(* IEC 61131-3 sources: daoli-st-library/DL_Algo (part 16) *)

(* ---- FB_DL_LoopCoupleDetect.st ---- *)
(*==============================================================================
 * 组件名称 (Component)  : FB_DL_LoopCoupleDetect
 * 所属子库 (Sublibrary) : DL_Algo
 * 当前版本 (Version)    : 1.0.1
 * 兼容性 (Platform)     : CODESYS 3.5+ / TwinCAT 3 / 汇川 InoProShop / 施耐德 Machine Expert
 *                         仅依赖 Standard.library（TON / R_TRIG），零厂商私有库
 * 功能描述 (Function)   : 回路耦合度在线探测。本回路上位激励期（bExcite 电平）
 *                         同步采集本回路 CV 增量 x 与邻回路 PV 增量 y，窗口内
 *                         计算皮尔逊互相关系数 r；|r| >= fCoupleThresh 且样本
 *                         充分 → bCoupled 锁存并输出耦合强度分级。为 Decouple2x2
 *                         提供投运判据（探测在先、解耦执行在后）。
 * 来源标签 (Origin)     : 自研线（IEC 61131-3 标准语义的道莅防御性实现，clean-room）
 * 分工声明 (Pairing)    : LoopCoupleDetect（探测，本件）↔ FB_DL_Decouple2x2
 *                         （解耦执行，既有件）：本件只输出耦合判据与强度分级，
 *                         不注入任何解耦补偿量、不修改解耦矩阵（R298 属主边界）；
 *                         与 FB_DL_CrossCorrelationDelay 分工：本件测「响应强度」
 *                         不测「延时幅值」，二者互补不重叠。
 * 边界语义 (Boundary)   : ① 相关系数除零防御：任一分母因子 <= eps → r 按 0
 *                         （邻回路无响应 = 无耦合语义，合法结果非故障）；
 *                         ② 非激励期（bExcite = FALSE）不采样不判据（判据串
 *                         相位因子，R281 口径）；
 *                         ③ 增量非有限拒收（NaN 自反 + Inf 差判）；
 *                         ④ 组态闸：窗深/阈值/最小样本 → 故障锁存。
 * 输出语义 (Fallback)   : 【R191】非激励期 → fCorrOut 保持末值、bCoupled 保持
 *                         锁存（耦合是资产属性，不随激励停而消失）；eFault 相
 *                         → 冻结 + bError = TRUE。
 * 码位     (Codes)      : 按 R297 范式零 16# 码位硬编码；错误出口 BOOL+ENUM(eCause)，
 *                         码位待主控收口统一派号。
 * 红线自检 (Redline)    : 7 项红线已自检：R1 零全局 ✓｜R2 零物理地址 ✓｜R3 纯 IEC ✓
 *                         R4 除零（双因子 eps 闸）/NaN 拒收/组态闸 ✓
 *                         R5 双语同行注释 ✓｜R6 CASE 带 ELSE 兜底迁 eFault ✓
 *                         R7 TON/R_TRIG 段 0 无条件刷新 ✓
 * 验收向量 (Acceptance) : V1 强耦合仿真（y = 0.8·x + 噪声）→ |r| ≈ 0.8+，
 *                         eStrength=eStrong，bCoupled=TRUE；
 *                         V2 独立回路（y 与 x 无关）→ |r| < 阈值，
 *                         eStrength=eNone；
 *                         V3 非激励期停止采样，样本数不增。
 * 修订历史 (Revision)   : 2026-11-20  v1.0.0  R49 首版（批 3 · 序号 13）
 *                        2026-11-20  v1.0.1  R51 文档级更正（R50 终审轻项）：3 处
 *                        相对指代禁词注释改为自含描述（R92/R68）；逻辑零变更
 *==============================================================================*)
TYPE E_DL_LcdStrength :
(
    eNone    := 0,                           (* 无耦合：|r| < 弱阈值 / No coupling *)
    eWeak    := 1,                           (* 弱耦合：|r| ∈ [弱阈, 强阈) / Weak coupling *)
    eStrong  := 2                            (* 强耦合：|r| >= 强阈值 / Strong coupling *)
);
END_TYPE

TYPE E_DL_LcdState :
(
    eIdle  := 0,                             (* 待使能 / Idle *)
    eProbe := 10,                            (* 激励探测运行 / Excitation probing *)
    eFault := 90                             (* 故障锁存相 / Fault latched phase *)
);
END_TYPE

TYPE E_DL_LcdCause :
(
    eNone       := 0,                        (* 无故障成因 / No cause *)
    eCfgIllegal := 1,                        (* 组态非法：窗深/阈值越域 / Illegal config *)
    ePhaseBad   := 2                         (* 非法相位兜底 / Illegal phase fallback *)
);
END_TYPE

FUNCTION_BLOCK FB_DL_LoopCoupleDetect
VAR_INPUT
    fCvThis   : LREAL := 0.0;                (* 本回路 CV 当前值（激励侧）[工程单位] / This loop CV value *)
    fPvNeighbor : LREAL := 0.0;              (* 邻回路 PV 当前值（响应侧）[工程单位] / Neighbor loop PV value *)
    bExcite   : BOOL := FALSE;               (* 本回路激励期电平（上位投运流程给出）[-] / Excitation period level *)
    nWinDepth : INT := 64;                   (* 互相关窗深，域 8..128 [点] / Correlation window depth *)
    fCoupleThresh : LREAL := 0.5;            (* 耦合判据阈值（|r| 门限），域 (0,1) [-] / Coupling threshold *)
    bEnable   : BOOL := TRUE;                (* 探测使能 [-] / Enable *)
    bReset    : BOOL := FALSE;               (* 复位命令，上升沿清窗与全部锁存 [-] / Reset command *)
END_VAR
VAR_OUTPUT
    fCorrOut  : LREAL;                       (* 当前窗口互相关系数 [-] / Window correlation coefficient *)
    eStrength : E_DL_LcdStrength;            (* 耦合强度分级出口（按最新窗口派生）[-] / Coupling strength outlet *)
    bCoupled  : BOOL;                        (* 耦合判据锁存位（复位沿清）[-] / Coupled latch *)
    nSampleCnt: INT;                         (* 窗口有效样本数 [点] / Valid sample count *)
    eState    : E_DL_LcdState;               (* 状态出口 / State outlet *)
    eCause    : E_DL_LcdCause;               (* 故障成因出口（R190 归因唯一） / Fault cause outlet *)
    bError    : BOOL;                        (* 故障锁存标志 [-] / Fault latch flag *)
END_VAR
VAR
    _eState  : E_DL_LcdState := E_DL_LcdState.eIdle;      (* 内部相位（CASE 唯一写入目标） / Internal phase *)
    _eCause  : E_DL_LcdCause := E_DL_LcdCause.eNone;      (* 故障成因锁存量 / Latched cause *)
    rtReset  : R_TRIG;                       (* 复位沿实例，段 0 无条件调用 / Reset edge instance *)
    _fCvPrev : LREAL;                        (* 上拍本回路 CV（增量基准）[工程单位] / Previous this-loop CV *)
    _fPvPrev : LREAL;                        (* 上拍邻回路 PV（增量基准）[工程单位] / Previous neighbor PV *)
    _aDx     : ARRAY[1..128] OF LREAL;       (* 本回路 CV 增量窗 [工程单位] / This-loop dCV window *)
    _aDy     : ARRAY[1..128] OF LREAL;       (* 邻回路 PV 增量窗 [工程单位] / Neighbor dPV window *)
    _nHead   : INT;                          (* 环形头游标 [-] / Ring head cursor *)
    _nFill   : INT;                          (* 窗填充数 [点] / Window fill count *)
    _nEff    : INT;                          (* 钳位后生效窗深 [点] / Clamped effective depth *)
    _fSumX   : LREAL;                        (* Σx [工程单位] / Sum x *)
    _fSumY   : LREAL;                        (* Σy [工程单位] / Sum y *)
    _fSumXY  : LREAL;                        (* Σxy [工程单位²] / Sum xy *)
    _fSumX2  : LREAL;                        (* Σx² [工程单位²] / Sum x2 *)
    _fSumY2  : LREAL;                        (* Σy² [工程单位²] / Sum y2 *)
    _fDen    : LREAL;                        (* 分母乘积（开方前）[-] / Denominator product *)
    _fR      : LREAL;                        (* 本拍相关系数 [-] / Correlation this scan *)
    _bFault  : BOOL;                         (* 故障锁存位 / Latched fault bit *)
    _bCfgBad : BOOL;                         (* 组态非法当拍量 / Illegal config this scan *)
    _i       : INT;                          (* 统计扫描游标（每趟重置，R227）[-] / Stats cursor *)
END_VAR
VAR CONSTANT
    DL_LCD_EPS  : LREAL := 1.0E-12;          (* 分母因子判零容差 [-] / Denominator epsilon *)
    DL_LCD_NMAX : INT   := 128;              (* 窗深容量上限 [点] / Window capacity limit *)
    DL_LCD_MIN  : INT   := 16;               (* 判据最小样本数（不足不判，防短窗误报）[点] / Min samples for verdict *)
    DL_LCD_WEAK : LREAL := 0.3;              (* 弱耦合门限（强度分级内界）[-] / Weak coupling bound *)
END_VAR

(* —— 段 0：当拍判据派生 + 实例无条件刷新（R228A） —— *)
_bCfgBad := (nWinDepth < 8) OR (nWinDepth > DL_LCD_NMAX) OR (fCoupleThresh <= 0.0) OR (fCoupleThresh >= 1.0);   (* 组态闸（R151 全引脚） / Config gate *)
rtReset(CLK := bReset);                      (* 复位沿每拍必调 / Reset edge every scan *)
_nEff := nWinDepth;                          (* 生效窗深初值 / Depth init *)
IF _nEff < 8 THEN
    _nEff := 8;                              (* 下限钳位 / Lower clamp *)
END_IF
IF _nEff > DL_LCD_NMAX THEN
    _nEff := DL_LCD_NMAX;                    (* 上限钳位（R308） / Upper clamp *)
END_IF

(* —— 段 1：单拍量预清零（R107） —— *)
_fSumX := 0.0;                               (* 累计量清零重算（每拍全路径派生，R285） / Sums recompute *)
_fSumY := 0.0;                               (* Σy 清零 / Sum y clear *)
_fSumXY := 0.0;                              (* Σxy 清零 / Sum xy clear *)
_fSumX2 := 0.0;                              (* Σx² 清零 / Sum x2 clear *)
_fSumY2 := 0.0;                              (* Σy² 清零 / Sum y2 clear *)
_fDen := 0.0;                                (* 分母清零（防残留触发除零） / Denominator clear *)
_fR := 0.0;                                  (* 相关系数缺省 0 / Correlation default *)

(* —— 段 2：复位沿处理（作用域：清故障 + 清窗 + 清锁存 + 基准重锚 + 迁 eIdle，R283 逐项声明） —— *)
IF rtReset.Q THEN
    _bFault := FALSE;                        (* 清故障锁存 / Clear fault *)
    _eCause := E_DL_LcdCause.eNone;          (* 清成因 / Clear cause *)
    _nFill := 0;                             (* 清窗填充 / Clear fill *)
    _nHead := 1;                             (* 头游标复位 / Head reset *)
    bCoupled := FALSE;                       (* 清耦合锁存 / Clear coupled latch *)
    fCorrOut := 0.0;                         (* 清相关系数出口 / Clear correlation outlet *)
    _fCvPrev := fCvThis;                     (* 增量基准重锚 / Re-anchor base *)
    _fPvPrev := fPvNeighbor;                 (* 邻回路 PV 增量基准重锚 / Re-anchor neighbor PV base *)
    _eState := E_DL_LcdState.eIdle;          (* 迁待机相 / Back to idle *)
END_IF

(* —— 段 3：组态闸故障锁存（R45 配对；锁存至复位沿，R189） —— *)
IF _bCfgBad AND NOT _bFault THEN
    _bFault := TRUE;                         (* 锁存故障位 / Latch fault *)
    _eCause := E_DL_LcdCause.eCfgIllegal;    (* 成因：组态非法 / Cause: illegal config *)
    _eState := E_DL_LcdState.eFault;         (* 同步迁故障相 / Migrate to fault *)
END_IF

(* —— 段 4：CASE 主状态机（ELSE 兜底迁 eFault，红线 6） —— *)
CASE _eState OF
    E_DL_LcdState.eIdle:                     (* 待机相：基准持续跟锚 / Idle *)
        _fCvPrev := fCvThis;                 (* 防待机期巨增量 / Anchor follow *)
        _fPvPrev := fPvNeighbor;             (* 邻回路 PV 基准持续跟锚（防待机期巨增量） / Neighbor PV base follow *)
        IF bEnable AND NOT _bFault THEN
            _eState := E_DL_LcdState.eProbe; (* 进入探测 / Enter probe *)
        END_IF
    E_DL_LcdState.eProbe:                    (* 探测相：仅激励期采样 + 窗口统计 / Probe *)
        IF NOT bEnable THEN
            _eState := E_DL_LcdState.eIdle;  (* 失能回待机 / Back to idle *)
        ELSE
            IF bExcite THEN                  (* 判据串相位因子：仅激励期采样（R281） / Sample only in excitation *)
                _aDx[_nHead] := fCvThis - _fCvPrev;       (* 本回路 CV 增量入窗 / This-loop dCV *)
                _aDy[_nHead] := fPvNeighbor - _fPvPrev;   (* 邻回路 PV 增量入窗 / Neighbor dPV *)
                IF (_aDx[_nHead] <> _aDx[_nHead]) OR (_aDy[_nHead] <> _aDy[_nHead])
                   OR ((_aDx[_nHead] - _aDx[_nHead]) <> (_aDx[_nHead] - _aDx[_nHead]))
                   OR ((_aDy[_nHead] - _aDy[_nHead]) <> (_aDy[_nHead] - _aDy[_nHead])) THEN
                    (* 非有限增量：不入统计不推进游标，基准照常跟锚 / Non-finite: skip *)
                    ;                        (* 空语句：ST 语法要求 THEN 分支非空，无副作用 / Empty statement, ST syntax requires non-empty branch *)
                ELSE
                    _nHead := _nHead + 1;    (* 有效样本：游标递进 / Head advance *)
                    IF _nHead > _nEff THEN
                        _nHead := 1;         (* 环回卷 / Ring wrap *)
                    END_IF
                    IF _nFill < _nEff THEN
                        _nFill := _nFill + 1;    (* 填充封顶 / Fill cap *)
                    END_IF
                END_IF
                _fCvPrev := fCvThis;         (* 基准推进 / Base advance *)
                _fPvPrev := fPvNeighbor;     (* 邻回路 PV 基准推进（与本拍采样配对） / Neighbor PV base advance *)
            END_IF
            _i := 1;                         (* 统计游标起头重置（R227） / Cursor reset *)
            WHILE _i <= _nFill DO            (* 逐点累计 / Per-point sums *)
                _fSumX := _fSumX + _aDx[_i]; (* Σx / Sum x *)
                _fSumY := _fSumY + _aDy[_i]; (* Σy / Sum y *)
                _fSumXY := _fSumXY + _aDx[_i] * _aDy[_i];   (* Σxy / Sum xy *)
                _fSumX2 := _fSumX2 + _aDx[_i] * _aDx[_i];   (* Σx² / Sum x2 *)
                _fSumY2 := _fSumY2 + _aDy[_i] * _aDy[_i];   (* Σy² / Sum y2 *)
                _i := _i + 1;                (* 游标递进 / Cursor advance *)
            END_WHILE
            IF _nFill >= 1 THEN
                _fDen := (DINT_TO_LREAL(_nFill) * _fSumX2 - _fSumX * _fSumX)
                       * (DINT_TO_LREAL(_nFill) * _fSumY2 - _fSumY * _fSumY);   (* 分母乘积（双因子联合闸） / Denominator product *)
            END_IF
            IF (_fDen > DL_LCD_EPS * DL_LCD_EPS) AND (_nFill >= 1) THEN
                _fR := (DINT_TO_LREAL(_nFill) * _fSumXY - _fSumX * _fSumY) / SQRT(_fDen);   (* 互相关 r：分母已过联合 eps 闸，无除零 / Correlation, denominator gated *)
                fCorrOut := _fR;             (* 相关系数出口更新（仅有效窗刷新） / Update outlet *)
                IF (_nFill >= DL_LCD_MIN) AND (_nFill * 10 >= 6 * _nEff) THEN
                    IF ABS(_fR) >= fCoupleThresh THEN
                        bCoupled := TRUE;    (* 耦合判据锁存至复位沿 / Coupled latch *)
                    END_IF
                    IF ABS(_fR) >= fCoupleThresh THEN
                        eStrength := E_DL_LcdStrength.eStrong;   (* 强耦合 / Strong *)
                    ELSIF ABS(_fR) >= DL_LCD_WEAK THEN
                        eStrength := E_DL_LcdStrength.eWeak;     (* 弱耦合 / Weak *)
                    ELSE
                        eStrength := E_DL_LcdStrength.eNone;     (* 无耦合（IF 链带 ELSE 兜底，R285） / None *)
                    END_IF
                END_IF
            END_IF
            nSampleCnt := _nFill;            (* 样本数出口镜像 / Sample count mirror *)
        END_IF
    E_DL_LcdState.eFault:                    (* 故障相：冻结保持，仅复位沿出 / Fault *)
        ;                                    (* 锁存回放（R28） / Replay from latch *)
    ELSE                                     (* 非法相位兜底迁安全态 / Illegal phase fallback *)
        _eState := E_DL_LcdState.eFault;     (* 迁故障相 / To fault *)
        _bFault := TRUE;                     (* 同步锁存 / Latch *)
        _eCause := E_DL_LcdCause.ePhaseBad;  (* 成因：非法相位 / Cause: illegal phase *)
END_CASE

(* —— 段 5：出口映射（bError/eState 同源，R191） —— *)
bError := _bFault;                           (* 故障标志镜像 / Fault flag mirror *)
eState := _eState;                           (* 状态出口 / State outlet *)
eCause := _eCause;                           (* 成因出口 / Cause outlet *)
END_FUNCTION_BLOCK

(* ---- FB_DL_LoopSignGuard.st ---- *)
(*==============================================================================
 * 组件名称 (Component)  : FB_DL_LoopSignGuard
 * 所属子库 (Sublibrary) : DL_Algo
 * 当前版本 (Version)    : 1.0.0
 * 兼容性 (Platform)     : CODESYS 3.5+ / TwinCAT 3 / 汇川 InoProShop / 施耐德 Machine Expert
 *                         仅依赖 Standard.library（TON），零厂商私有库
 * 功能描述 (Function)   : 回路正反作用符号在线自检（调试期防呆）。以增量对
 *                         (dCV, dPV) 为样本，窗口内计算皮尔逊相关系数
 *                         r = (nΣxy - ΣxΣy) / sqrt((nΣx²-(Σx)²)·(nΣy²-(Σy)²))：
 *                         r > fSignThresh → 判正向作用（CV 增大 PV 随之增大）；
 *                         r < -fSignThresh → 判反向作用；|r| 不足 → 未定。
 *                         期望作用 eExpect 与实测作用不一致 → bSignSuspect
 *                         锁存（接线反接/正反作用组态错防呆）。
 * 来源标签 (Origin)     : 自研线（IEC 61131-3 标准语义的道莅防御性实现，clean-room）
 * 边界语义 (Boundary)   : ① 相关系数除零防御：分母任一因子 <= eps（窗口内
 *                         CV 或 PV 无变化，如手动手假输入）→ r 按 0 处理（未定），
 *                         不产生 Inf/NaN；
 *                         ② 样本拒收：dCV/dPV 非有限（NaN/Inf 差判）不入窗；
 *                         ③ 判据串相位因子：仅 nSample >= 窗深 60% 后才判
 *                         （样本不足不判，防启动段误报，R281 口径）；
 *                         ④ 组态闸：窗深 < 8 / 阈值域 (0,1) 外 → 故障。
 * 输出语义 (Fallback)   : 【R191】样本不足期 → eSignOut = eUnknown，bSignSuspect
 *                         保持 FALSE；eFault 相 → 判据输出冻结保持末值。
 * 码位     (Codes)      : 按 R297 范式零 16# 码位硬编码；错误出口 BOOL+ENUM(eCause)，
 *                         码位待主控收口统一派号。
 * 红线自检 (Redline)    : 7 项红线已自检：R1 零全局 ✓｜R2 零物理地址 ✓｜R3 纯 IEC ✓
 *                         R4 除零（双因子 eps 闸）/NaN 拒收/组态闸 ✓
 *                         R5 双语同行注释 ✓｜R6 CASE 带 ELSE 兜底迁 eFault ✓
 *                         R7 TON/R_TRIG 段 0 无条件刷新 ✓
 * 验收向量 (Acceptance) : V1 同向增量样本 32 点 → r≈1 → eSignOut=eDirect；
 *                         V2 反向增量样本 → r≈-1 → eSignOut=eReverse，若
 *                         eExpect=eDirect → bSignSuspect=TRUE；
 *                         V3 恒定 PV（分母 0）→ eSignOut=eUnknown，不误报。
 * 修订历史 (Revision)   : 2026-11-20  v1.0.0  R49 首版（批 3 · 序号 11）
 *==============================================================================*)
TYPE E_DL_LsgSign :
(
    eUnknown := 0,                           (* 未定（样本不足或相关性弱） / Unknown *)
    eDirect  := 1,                           (* 正向作用：CV↑ → PV↑ / Direct acting *)
    eReverse := 2                            (* 反向作用：CV↑ → PV↓ / Reverse acting *)
);
END_TYPE

TYPE E_DL_LsgState :
(
    eIdle  := 0,                             (* 待使能 / Idle *)
    eLearn := 10,                            (* 增量样本采集学习中 / Learning *)
    eFault := 90                             (* 故障锁存相 / Fault latched phase *)
);
END_TYPE

TYPE E_DL_LsgCause :
(
    eNone       := 0,                        (* 无故障成因 / No cause *)
    eCfgIllegal := 1,                        (* 组态非法：窗深/阈值越域 / Illegal config *)
    ePhaseBad   := 2                         (* 非法相位兜底 / Illegal phase fallback *)
);
END_TYPE

FUNCTION_BLOCK FB_DL_LoopSignGuard
VAR_INPUT
    fCvNow    : LREAL := 0.0;                (* 控制量当前值（CV）[工程单位] / CV current value *)
    fPvNow    : LREAL := 0.0;                (* 过程量当前值（PV）[工程单位] / PV current value *)
    nWinDepth : INT := 32;                   (* 增量样本窗深，域 8..64 [点] / Sample window depth *)
    fSignThresh : LREAL := 0.6;              (* 判向阈值（|r| 门限），域 (0.0, 1.0) [-] / Sign verdict threshold *)
    eExpect   : E_DL_LsgSign := E_DL_LsgSign.eDirect;   (* 期望作用方向（组态声明）[-] / Expected acting direction *)
    bEnable   : BOOL := TRUE;                (* 自检使能 [-] / Enable *)
    bReset    : BOOL := FALSE;               (* 复位命令，上升沿清全部样本与锁存 [-] / Reset command *)
END_VAR
VAR_OUTPUT
    eSignOut     : E_DL_LsgSign;             (* 实测作用方向出口 / Measured sign outlet *)
    fCorrCoef    : LREAL;                    (* 当前窗口皮尔逊相关系数 [-] / Pearson correlation of window *)
    nSampleCnt   : INT;                      (* 窗口内有效样本数 [点] / Valid sample count *)
    bSignSuspect : BOOL;                     (* 作用方向与期望不符锁存位（复位沿清）[-] / Sign-suspect latch *)
    eState       : E_DL_LsgState;            (* 状态出口 / State outlet *)
    eCause       : E_DL_LsgCause;            (* 故障成因出口（R190 归因唯一） / Fault cause outlet *)
    bError       : BOOL;                     (* 故障锁存标志 [-] / Fault latch flag *)
END_VAR
VAR
    _eState  : E_DL_LsgState := E_DL_LsgState.eIdle;      (* 内部相位（CASE 唯一写入目标） / Internal phase *)
    _eCause  : E_DL_LsgCause := E_DL_LsgCause.eNone;      (* 故障成因锁存量 / Latched cause *)
    rtReset  : R_TRIG;                       (* 复位沿实例，段 0 无条件调用 / Reset edge instance *)
    _fCvPrev : LREAL;                        (* 上拍 CV（增量基准）[工程单位] / Previous CV *)
    _fPvPrev : LREAL;                        (* 上拍 PV（增量基准）[工程单位] / Previous PV *)
    _aDx     : ARRAY[1..64] OF LREAL;        (* dCV 样本窗 [工程单位] / dCV window *)
    _aDy     : ARRAY[1..64] OF LREAL;        (* dPV 样本窗 [工程单位] / dPV window *)
    _nHead   : INT;                          (* 环形头游标 [-] / Ring head cursor *)
    _nFill   : INT;                          (* 窗口填充数 [点] / Window fill count *)
    _nEff    : INT;                          (* 钳位后生效窗深 [点] / Clamped effective depth *)
    _fSumX   : LREAL;                        (* Σx 累计 [工程单位] / Sum x *)
    _fSumY   : LREAL;                        (* Σy 累计 [工程单位] / Sum y *)
    _fSumXY  : LREAL;                        (* Σxy 累计 [工程单位²] / Sum xy *)
    _fSumX2  : LREAL;                        (* Σx² 累计 [工程单位²] / Sum x2 *)
    _fSumY2  : LREAL;                        (* Σy² 累计 [工程单位²] / Sum y2 *)
    _fDenX   : LREAL;                        (* 分母因子 1：nΣx²-(Σx)² [-] / Denominator factor 1 *)
    _fDenY   : LREAL;                        (* 分母因子 2：nΣy²-(Σy)² [-] / Denominator factor 2 *)
    _fDen    : LREAL;                        (* 相关系数分母（开方前乘积）[-] / Correlation denominator *)
    _fR      : LREAL;                        (* 本拍相关系数 [-] / Correlation this scan *)
    _eSign   : E_DL_LsgSign := E_DL_LsgSign.eUnknown;     (* 实测方向锁存 / Measured sign latch *)
    _bFault  : BOOL;                         (* 故障锁存位 / Latched fault bit *)
    _bCfgBad : BOOL;                         (* 组态非法当拍量 / Illegal config this scan *)
    _i       : INT;                          (* 统计扫描游标（每趟重置，R227）[-] / Stats cursor *)
END_VAR
VAR CONSTANT
    DL_LSG_EPS   : LREAL := 1.0E-12;         (* 分母因子判零容差 [-] / Denominator epsilon *)
    DL_LSG_NMAX  : INT   := 64;              (* 窗深容量上限 [点] / Window capacity limit *)
END_VAR

(* —— 段 0：当拍判据派生 + 实例无条件刷新（R228A） —— *)
_bCfgBad := (nWinDepth < 8) OR (nWinDepth > DL_LSG_NMAX) OR (fSignThresh <= 0.0) OR (fSignThresh >= 1.0);   (* 组态闸（R151 全引脚） / Config gate *)
rtReset(CLK := bReset);                      (* 复位沿每拍必调 / Reset edge every scan *)
_nEff := nWinDepth;                          (* 生效窗深初值 / Effective depth init *)
IF _nEff < 8 THEN
    _nEff := 8;                              (* 窗深下限钳位 / Depth lower clamp *)
END_IF
IF _nEff > DL_LSG_NMAX THEN
    _nEff := DL_LSG_NMAX;                    (* 窗深上限钳位（R308） / Depth upper clamp *)
END_IF

(* —— 段 1：单拍量预清零（R107） —— *)
_fSumX := 0.0;                               (* 累计量清零重算（每拍全路径派生，R285） / Sums recompute *)
_fSumY := 0.0;                               (* Σy 清零 / Sum y clear *)
_fSumXY := 0.0;                              (* Σxy 清零 / Sum xy clear *)
_fSumX2 := 0.0;                              (* Σx² 清零 / Sum x2 clear *)
_fSumY2 := 0.0;                              (* Σy² 清零 / Sum y2 clear *)
_fDen := 0.0;                                (* 分母清零（防 _nFill=0 残留触发除零） / Denominator clear *)
_fR := 0.0;                                  (* 相关系数缺省 0（未定语义） / Correlation default zero *)

(* —— 段 2：复位沿处理（作用域：清故障 + 清窗 + 清方向锁存 + 清嫌疑锁存 + 迁 eIdle，R283 逐项声明） —— *)
IF rtReset.Q THEN
    _bFault := FALSE;                        (* 清故障锁存 / Clear fault *)
    _eCause := E_DL_LsgCause.eNone;          (* 清成因 / Clear cause *)
    _nFill := 0;                             (* 清窗填充 / Clear fill *)
    _nHead := 1;                             (* 头游标复位 / Head reset *)
    _eSign := E_DL_LsgSign.eUnknown;         (* 方向回未定 / Sign back to unknown *)
    bSignSuspect := FALSE;                   (* 清嫌疑锁存 / Clear suspect latch *)
    _fCvPrev := fCvNow;                      (* 增量基准重锚（防复位后巨增量） / Re-anchor increment base *)
    _fPvPrev := fPvNow;                      (* 同前一项，基准跟锚 / Same as previous line, anchor follow *)
    _eState := E_DL_LsgState.eIdle;          (* 迁待机相 / Back to idle *)
END_IF

(* —— 段 3：组态闸故障锁存（R45 配对；锁存至复位沿，R189） —— *)
IF _bCfgBad AND NOT _bFault THEN
    _bFault := TRUE;                         (* 锁存故障位 / Latch fault *)
    _eCause := E_DL_LsgCause.eCfgIllegal;    (* 成因：组态非法 / Cause: illegal config *)
    _eState := E_DL_LsgState.eFault;         (* 同步迁故障相 / Migrate to fault *)
END_IF

(* —— 段 4：CASE 主状态机（ELSE 兜底迁 eFault，红线 6） —— *)
CASE _eState OF
    E_DL_LsgState.eIdle:                     (* 待机相 / Idle *)
        _fCvPrev := fCvNow;                  (* 增量基准持续跟锚（防待机期累积巨增量） / Anchor follow *)
        _fPvPrev := fPvNow;                  (* 同前一项，基准跟锚 / Same as previous line, anchor follow *)
        IF bEnable AND NOT _bFault THEN
            _eState := E_DL_LsgState.eLearn; (* 进入学习 / Enter learn *)
        END_IF
    E_DL_LsgState.eLearn:                    (* 学习相：增量采样 + 窗口统计 / Learn *)
        IF NOT bEnable THEN
            _eState := E_DL_LsgState.eIdle;  (* 失能回待机 / Back to idle *)
        ELSE
            _aDx[_nHead] := fCvNow - _fCvPrev;   (* dCV 增量入窗 / dCV into window *)
            _aDy[_nHead] := fPvNow - _fPvPrev;   (* dPV 增量入窗 / dPV into window *)
            IF (_aDx[_nHead] <> _aDx[_nHead]) OR (_aDy[_nHead] <> _aDy[_nHead])
               OR ((_aDx[_nHead] - _aDx[_nHead]) <> (_aDx[_nHead] - _aDx[_nHead]))
               OR ((_aDy[_nHead] - _aDy[_nHead]) <> (_aDy[_nHead] - _aDy[_nHead])) THEN
                (* 非有限增量：不入统计、不推进游标，基准照常跟锚（NaN 拒收口径） / Non-finite: skip, anchor follows *)
                _fCvPrev := fCvNow;          (* 基准照常跟锚 / Anchor follow *)
                _fPvPrev := fPvNow;          (* 同前一项，基准跟锚 / Same as previous line, anchor follow *)
            ELSE
                _nHead := _nHead + 1;        (* 有效样本：头游标递进 / Head advance *)
                IF _nHead > _nEff THEN
                    _nHead := 1;             (* 环回卷（下标先判后增） / Ring wrap *)
                END_IF
                IF _nFill < _nEff THEN
                    _nFill := _nFill + 1;    (* 填充计数封顶 / Fill cap *)
                END_IF
                _fCvPrev := fCvNow;          (* 基准推进 / Base advance *)
                _fPvPrev := fPvNow;          (* 同前一项，基准跟锚 / Same as previous line, anchor follow *)
            END_IF
            _i := 1;                         (* 统计游标起头重置（R227） / Cursor reset *)
            WHILE _i <= _nFill DO            (* 逐点累计（窗口内下标已钳位） / Per-point sums *)
                _fSumX := _fSumX + _aDx[_i]; (* Σx / Sum x *)
                _fSumY := _fSumY + _aDy[_i]; (* Σy / Sum y *)
                _fSumXY := _fSumXY + _aDx[_i] * _aDy[_i];   (* Σxy / Sum xy *)
                _fSumX2 := _fSumX2 + _aDx[_i] * _aDx[_i];   (* Σx² / Sum x2 *)
                _fSumY2 := _fSumY2 + _aDy[_i] * _aDy[_i];   (* Σy² / Sum y2 *)
                _i := _i + 1;                (* 游标递进 / Cursor advance *)
            END_WHILE
            IF _nFill >= 1 THEN
                _fDenX := DINT_TO_LREAL(_nFill) * _fSumX2 - _fSumX * _fSumX;   (* 分母因子 1 / Denominator factor 1 *)
                _fDenY := DINT_TO_LREAL(_nFill) * _fSumY2 - _fSumY * _fSumY;   (* 分母因子 2 / Denominator factor 2 *)
                _fDen := _fDenX * _fDenY;    (* 开方前乘积 / Product before sqrt *)
            END_IF
            IF (_fDen > DL_LSG_EPS * DL_LSG_EPS) AND (_nFill >= 1) THEN
                _fR := (DINT_TO_LREAL(_nFill) * _fSumXY - _fSumX * _fSumY) / SQRT(_fDen);   (* 皮尔逊 r：分母已过乘积 eps 闸（乘积闸等价双因子闸），无除零 / Pearson r, denominator gated *)
                IF _fR > fSignThresh THEN
                    _eSign := E_DL_LsgSign.eDirect;      (* 判正向 / Direct *)
                ELSIF _fR < (-fSignThresh) THEN
                    _eSign := E_DL_LsgSign.eReverse;     (* 判反向 / Reverse *)
                ELSE
                    _eSign := E_DL_LsgSign.eUnknown;     (* 相关性弱：未定（IF 链带 ELSE 兜底，R285） / Weak: unknown *)
                END_IF
            ELSE
                _eSign := E_DL_LsgSign.eUnknown;         (* 窗内无变化/无样本：未定（边界①） / Degenerate: unknown *)
            END_IF
            fCorrCoef := _fR;                (* 相关系数出口镜像 / Correlation mirror *)
            nSampleCnt := _nFill;            (* 样本数出口镜像 / Sample count mirror *)
            eSignOut := _eSign;              (* 方向出口镜像 / Sign mirror *)
            IF (_nFill * 10 >= 6 * _nEff) THEN
                (* 判据串相位因子：填充 >= 60% 才比对期望（R281 口径，整数交叉乘比避免浮点除） / Verdict gated at 60% fill, integer cross-multiply *)
                IF (_eSign = E_DL_LsgSign.eDirect OR _eSign = E_DL_LsgSign.eReverse)
                   AND (_eSign <> eExpect) THEN
                    bSignSuspect := TRUE;    (* 方向与期望不符：嫌疑锁存至复位沿 / Suspect latch *)
                END_IF
            END_IF
        END_IF
    E_DL_LsgState.eFault:                    (* 故障相：冻结保持，仅复位沿出 / Fault *)
        ;                                    (* 锁存回放（R28） / Replay from latch *)
    ELSE                                     (* 非法相位兜底迁安全态 / Illegal phase fallback *)
        _eState := E_DL_LsgState.eFault;     (* 迁故障相 / To fault *)
        _bFault := TRUE;                     (* 同步锁存 / Latch *)
        _eCause := E_DL_LsgCause.ePhaseBad;  (* 成因：非法相位 / Cause: illegal phase *)
END_CASE

(* —— 段 5：出口映射（bError/eState 同源，R191） —— *)
bError := _bFault;                           (* 故障标志镜像 / Fault flag mirror *)
eState := _eState;                           (* 状态出口 / State outlet *)
eCause := _eCause;                           (* 成因出口 / Cause outlet *)
END_FUNCTION_BLOCK

(* ---- FB_DL_LoopWaveInject.st ---- *)
(*==============================================================================
 * 组件名称 (Component)  : FB_DL_LoopWaveInject
 * 所属子库 (Sublibrary) : DL_Algo
 * 当前版本 (Version)    : 1.0.0
 * 兼容性 (Platform)     : CODESYS 3.5 / TwinCAT 3 / 汇川 InoProShop / Machine Expert
 *                         仅依赖纯 IEC 61131-3 标准元素，零厂商方言
 * 功能描述 (Function)   : PID 回路调试激励源：正弦/方波/阶跃三型可选，输出经
 *                         委托 FB_DL_RateLimiter 斜率保护后叠加到给定值。
 *                         相位累加器按采样周期推进（周期越界钳制）；
 *                         使能撤销后目标平滑归零（经限速器自然回零），
 *                         完全禁用期间输出冻结 0，不塞伪值。
 * 溯源 (Origin)         : 道莅 clean-room 防御性实现
 * 本文件内含 (Contains) : TYPE E_DL_WaveType / TYPE E_DL_InjErr /
 *                         FUNCTION_BLOCK FB_DL_LoopWaveInject
 * 依赖 (Depends)        : DL_Algo/FB_DL_RateLimiter、DL_MathData/FC_DL_TimeToLrealSec
 * 红线自检 (Redline)    : 无外部全局变量、无硬件地址直引 ｜ 全变量中英双语同行注释
 *                         防除零 + 量程钳位 + 非有限值防御 ｜ 枚举成员全部显式赋值
 *                         委托限速器实例每周期无条件调用（仅输入条件化）｜
 *                         相位累加器每周期无条件刷新 ｜ CASE 含 ELSE 兜底
 * 错误码表 (Codes)      : 16#0002_3710 就绪
 *                         16#0002_3711 信息级 幅值越界(已钳制)
 *                         16#0002_3712 信息级 周期非法(已钳制)
 *                         16#0002_3713 信息级 斜率限制非法(已钳制)
 *                         16#0002_3714 信息级 注入激活中
 * 修订历史 (Revision)   : 2026-11-17  v1.0.0  首版入库 · R27 · 阶段三批 1
 * 验收向量 (Acceptance) : SIN 幅 10% 周期 10 s → 输出 5 Hz 采样下按 2*pi*相位 正弦；
 *                         幅值 120 → 钳 100 且 3711；周期 0 → 钳下限且 3712；
 *                         bEnable 撤销 → 输出按斜率回零后冻结 0
 *============================================================================*)

(*-----------------------------------------------------------------------------
 * 枚举: E_DL_WaveType（归属 DL_Algo，波形类型）
 *----------------------------------------------------------------------------*)
TYPE E_DL_WaveType :
(
    eWaveSin  := 0,    // 正弦波 / Sine wave
    eWaveSqr  := 1,    // 方波（半周期正半幅，半周期负半幅）/ Square wave
    eWaveStep := 2     // 阶跃（激活期间恒幅）/ Step wave
);
END_TYPE

(*-----------------------------------------------------------------------------
 * 枚举: E_DL_InjErr（归属 DL_Algo，与 FB_DL_LoopWaveInject 同文件）
 *----------------------------------------------------------------------------*)
TYPE E_DL_InjErr :
(
    eReady      := 16#0002_3710,    // 就绪 / Ready
    eAmpClamped := 16#0002_3711,    // 信息级：幅值越界已钳制 / Info: amplitude clamped
    ePeriodBad  := 16#0002_3712,    // 信息级：周期非法已钳制 / Info: period clamped
    eSlewBad    := 16#0002_3713,    // 信息级：斜率限制非法已钳制 / Info: slew limit clamped
    eActive     := 16#0002_3714     // 信息级：注入激活中 / Info: injection active
);
END_TYPE

(*==============================================================================
 * 功能块: FB_DL_LoopWaveInject
 * 调用约定: 每个扫描周期无条件调用一次；tSampleTime 必须注入真实任务间隔。
 *============================================================================*)
FUNCTION_BLOCK FB_DL_LoopWaveInject
VAR_INPUT
    bEnable      : BOOL;               // 注入使能 / Injection enable
    eWaveType    : E_DL_WaveType;      // 波形类型 SIN/SQR/STEP / Wave type selection
    fAmplitude   : REAL;               // 幅值 [百分数]，有效域 0~100 / Amplitude [percent]
    fPeriod_s    : REAL;               // 周期 [秒]，有效域 0.1~600 / Period [s]
    fSlewLimit   : REAL;               // 斜率限制 [百分数每秒]，有效域 0.01~100 / Slew limit [percent per s]
    tSampleTime  : TIME := T#100MS;    // 采样周期，调用方注入真实任务间隔 / Sample period, caller-injected task interval
END_VAR
VAR_OUTPUT
    fInjectOut   : REAL;               // 注入量 [百分数] / Injection output [percent]
    bActive      : BOOL;               // 注入有效（输出非零或正在回零）/ Injection active flag
    eErr         : E_DL_InjErr;        // 错误码 / Error code
END_VAR
VAR
    fbLimiter    : FB_DL_RateLimiter;  // 委托限速器实例（每周期无条件调用）/ Delegate rate limiter instance
    fPhase       : REAL;               // 相位累加器 [0~1)，无量纲 / Phase accumulator [0..1)
    fAmpUse      : REAL;               // 生效幅值（钳位后）[百分数] / Effective amplitude [percent]
    fPeriodUse   : REAL;               // 生效周期（钳位后）[秒] / Effective period [s]
    fSlewUse     : REAL;               // 生效斜率（钳位后）[百分数每秒] / Effective slew limit [percent per s]
    fDtSec       : LREAL;              // 采样周期秒值（委托换算）[秒] / Sample period in seconds via delegate
    fWaveTarget  : REAL;               // 波形目标值（限速器输入）[百分数] / Wave target value, limiter input [percent]
    fTwoPi       : REAL := 6.283185307179586;   // 圆周率二倍 [弧度] / Two pi [rad]
    bLimErr      : BOOL;               // 委托限速器故障位 / Delegate rate limiter fault bit
END_VAR
VAR CONSTANT
    DL_INJ_AMP_MIN    : REAL := 0.0;    // 幅值下限 [百分数] / Amplitude lower bound [percent]
    DL_INJ_AMP_MAX    : REAL := 100.0;  // 幅值上限 [百分数] / Amplitude upper bound [percent]
    DL_INJ_PERIOD_MIN : REAL := 0.1;    // 周期下限 [秒] / Period lower bound [s]
    DL_INJ_PERIOD_MAX : REAL := 600.0;  // 周期上限 [秒] / Period upper bound [s]
    DL_INJ_SLEW_MIN   : REAL := 0.01;   // 斜率下限 [百分数每秒] / Slew lower bound [percent per s]
    DL_INJ_SLEW_MAX   : REAL := 100.0;  // 斜率上限 [百分数每秒] / Slew upper bound [percent per s]
    DL_INJ_INF_MAX    : REAL := 1.0E30; // 非有限值判定幅值上限 / Magnitude bound for finite-value check
    DL_INJ_ZERO       : REAL := 0.0;    // 零值常量，避免裸字面量 / Zero constant
    DL_INJ_TOL        : REAL := 1.0E-6; // 浮点比较容差 / Float comparison tolerance
END_VAR

(*------------------------------------------------------------------------------
 * 段 1｜委托限速器每周期无条件调用（仅输入条件化）：斜率保护永不断流
 *----------------------------------------------------------------------------*)
fbLimiter(bEnable := TRUE,                    // 限速器自身常开，方向限速由 fRate 引脚承载 / limiter always enabled
          fIn := fWaveTarget,                 // 波形目标作为限速输入 / wave target as limiter input
          fRateUp := fSlewUse,                // 上升斜率限制 [百分数每秒] / rising slew limit
          fRateDown := fSlewUse,              // 下降斜率限制（回零同样受保护）/ falling slew limit
          bTrack := FALSE,                    // 不使用跟踪回投 / no tracking
          fTrackValue := DL_INJ_ZERO,         // 跟踪值未用 / track value unused
          tSampleTime := tSampleTime,         // 采样周期透传 / sample period passed through
          fOut => fInjectOut,                 // 限速输出直接对外 / rate-limited output exported
          bError => bLimErr);                 // 委托故障位回收 / delegate fault bit captured

(*------------------------------------------------------------------------------
 * 段 2｜非有限值与参数钳位：越界钳制并置信息码（先到先得，斜率最后判）
 *----------------------------------------------------------------------------*)
IF (fAmplitude <> fAmplitude) OR (ABS(fAmplitude) > DL_INJ_INF_MAX) THEN
    fAmpUse := DL_INJ_AMP_MAX;                       // 非有限幅值按上限处置 / non-finite amplitude treated as upper bound
    eErr := E_DL_InjErr.eAmpClamped;                 // 信息级：幅值越界 / info: amplitude clamped
ELSIF fAmplitude < DL_INJ_AMP_MIN THEN
    fAmpUse := DL_INJ_AMP_MIN;                       // 下限钳位 / floored
    eErr := E_DL_InjErr.eAmpClamped;                 // 信息级：幅值越界 / info: amplitude clamped
ELSIF fAmplitude > DL_INJ_AMP_MAX THEN
    fAmpUse := DL_INJ_AMP_MAX;                       // 上限钳位 / capped
    eErr := E_DL_InjErr.eAmpClamped;                 // 信息级：幅值越界 / info: amplitude clamped
ELSE
    fAmpUse := fAmplitude;                           // 幅值域内 / amplitude in range
END_IF
IF (fPeriod_s <> fPeriod_s) OR (ABS(fPeriod_s) > DL_INJ_INF_MAX) THEN
    fPeriodUse := DL_INJ_PERIOD_MIN;                 // 非有限周期按下限处置（防除零）/ non-finite period treated as lower bound
    IF eErr = E_DL_InjErr.eReady THEN
        eErr := E_DL_InjErr.ePeriodBad;              // 信息级：周期非法 / info: period clamped
    END_IF
ELSIF fPeriod_s < DL_INJ_PERIOD_MIN THEN
    fPeriodUse := DL_INJ_PERIOD_MIN;                 // 周期下限钳位（防除零）/ period floored
    IF eErr = E_DL_InjErr.eReady THEN
        eErr := E_DL_InjErr.ePeriodBad;              // 信息级：周期非法 / info: period clamped
    END_IF
ELSIF fPeriod_s > DL_INJ_PERIOD_MAX THEN
    fPeriodUse := DL_INJ_PERIOD_MAX;                 // 周期上限钳位 / period capped
    IF eErr = E_DL_InjErr.eReady THEN
        eErr := E_DL_InjErr.ePeriodBad;              // 信息级：周期非法 / info: period clamped
    END_IF
ELSE
    fPeriodUse := fPeriod_s;                         // 周期域内 / period in range
END_IF
IF (fSlewLimit <> fSlewLimit) OR (ABS(fSlewLimit) > DL_INJ_INF_MAX) THEN
    fSlewUse := DL_INJ_SLEW_MAX;                     // 非有限斜率按上限处置 / non-finite slew treated as upper bound
    IF eErr = E_DL_InjErr.eReady THEN
        eErr := E_DL_InjErr.eSlewBad;                // 信息级：斜率非法 / info: slew clamped
    END_IF
ELSIF (fSlewLimit < DL_INJ_SLEW_MIN) OR (fSlewLimit > DL_INJ_SLEW_MAX) THEN
    IF fSlewLimit < DL_INJ_SLEW_MIN THEN
        fSlewUse := DL_INJ_SLEW_MIN;                 // 斜率下限钳位 / slew floored
    ELSE
        fSlewUse := DL_INJ_SLEW_MAX;                 // 斜率上限钳位 / slew capped
    END_IF
    IF eErr = E_DL_InjErr.eReady THEN
        eErr := E_DL_InjErr.eSlewBad;                // 信息级：斜率非法 / info: slew clamped
    END_IF
ELSE
    fSlewUse := fSlewLimit;                          // 斜率域内 / slew in range
END_IF

(*------------------------------------------------------------------------------
 * 段 3｜采样周期委托换算（FC_DL_TimeToLrealSec）与除零防御
 *----------------------------------------------------------------------------*)
fDtSec := FC_DL_TimeToLrealSec(tIn := tSampleTime);  // 采样周期秒值（委托换算）/ sample period in seconds via delegate
IF (fDtSec <> fDtSec) OR (fDtSec < DL_INJ_TOL) OR (fDtSec > REAL_TO_LREAL(DL_INJ_INF_MAX)) THEN
    fDtSec := LREAL#0.1;                             // 非法采样周期按 0.1 s 兜底（防除零）/ illegal sample period falls back to 0.1 s
END_IF

(*------------------------------------------------------------------------------
 * 段 4｜相位累加器：每周期无条件推进，按波形周期归一化回卷
 *----------------------------------------------------------------------------*)
IF bEnable THEN
    fPhase := fPhase + LREAL_TO_REAL(fDtSec / REAL_TO_LREAL(fPeriodUse));   // 相位推进 [无量纲] / phase advance
    WHILE fPhase >= 1.0 DO
        fPhase := fPhase - 1.0;                      // 相位回卷 [0~1) / phase wrap into [0..1)
    END_WHILE
END_IF

(*------------------------------------------------------------------------------
 * 段 5｜波形目标计算：CASE 含 ELSE 兜底（默认目标 0）
 *----------------------------------------------------------------------------*)
IF bEnable THEN
    CASE eWaveType OF
        E_DL_WaveType.eWaveSin:
            fWaveTarget := fAmpUse * SIN(fPhase * fTwoPi);          // 正弦目标 [百分数] / sine target [percent]
        E_DL_WaveType.eWaveSqr:
            IF fPhase < 0.5 THEN
                fWaveTarget := fAmpUse;                             // 方波正半幅 [百分数] / square positive half [percent]
            ELSE
                fWaveTarget := -fAmpUse;                            // 方波负半幅 [百分数] / square negative half [percent]
            END_IF
        E_DL_WaveType.eWaveStep:
            fWaveTarget := fAmpUse;                                 // 阶跃恒幅目标 [百分数] / step target [percent]
        ELSE
            fWaveTarget := DL_INJ_ZERO;                             // 非法波形兜底目标 0 / illegal wave type, target zero
    END_CASE
    bActive := TRUE;                                 // 注入激活 / injection active
    IF eErr = E_DL_InjErr.eReady THEN
        eErr := E_DL_InjErr.eActive;                 // 信息级：注入激活中 / info: injection active
    END_IF
ELSE
    fWaveTarget := DL_INJ_ZERO;                      // 禁用目标 0（经限速器平滑回零）/ disabled target zero, slews down
    bActive := ABS(fInjectOut) > DL_INJ_TOL;         // 回零期间仍视为激活 / active while settling to zero
    IF ABS(fInjectOut) <= DL_INJ_TOL THEN
        fInjectOut := DL_INJ_ZERO;                   // 回零完成冻结 0（禁用期不塞伪值）/ settled frozen at zero
        bActive := FALSE;                            // 注入失效 / injection inactive
        fPhase := DL_INJ_ZERO;                       // 相位复位（下次启用从零相位起）/ phase reset for next enable
    END_IF
END_IF
END_FUNCTION_BLOCK

(* ---- FB_DL_LossInWeightFeeder.st ---- *)
(*
  ==================================================================
  组件名 Component  : FB_DL_LossInWeightFeeder
  分类   Category   : DL_Algo
  复杂度 Complexity  : cx5
  版本   Version    : 1.0.1
  功能   Purpose    : 失重式给料控制。称重 w(t) 一阶差分求失重速率（负变化为正
                      给料率），一阶低通滤波后进 PI 闭环调节螺旋输出；低料位触发
                      补料相（输出冻结归零、计量与速率估计暂停），补料完成沿或
                      超时退出；批量累计达目标判批次结束。速率长期为零而输出非零
                      判 eNoLossRate；称重突跳超物理限判 eWeightNoise。
  来源   Source     : t2-2-lbp（与 FB_DL_BatchDosingControl 分工：连续失重 vs 批次定量）
  溯源   Origin     : IEC 61131-3 标准语义的道莅防御性实现；失重秤连续给料为公开
                      工艺语义，clean-room 自研实现，未复制任何闭源代码行。
  平台   Platform   : 纯 IEC 61131-3（TON / R_TRIG / LREAL，无私有库）
  作者   Author     : 道莅代码库 · PLC 编程专家（R56）
  ------------------------------------------------------------------
  同拍双窗配比约束（R100）：tRefillTo（补料超时窗）与 tNoRateTo（无速率确认窗）
                      职责分离、分属不同相，IN 串各自相位闸，无同拍并跑；
                      配比约束 tRefillTo > tNoRateTo 在组态域闸内判故障。
  边界 Boundary     :
                      一 本件只算给料输出与批量累计，不驱动螺旋电机本体、不控补料阀
                         （补料阀由外部按 bRefilling 执行，属主边界）；
                      二 失重速率方向约定：w(t) 递减 = 给料，速率为正；
                      三 补料相冻结语义（R191 显式声明）：输出归零、累计与速率估计
                         全部暂停，恢复后从冻结点继续；
                      四 相级看门狗使能只用相驻留本身（R145）；
                      五 故障锁存解除路径 = bReset 上升沿（唯一路径，R188）；
                      六 无全局变量、无外部变量声明、无物理地址寻址。
  输出契约 Output contract:
                      fRateOut 为 PI 后给料输出（0..fOutMax）；bDosing / bRefilling
                      为相位派生电平；fBatchAcc 为批量累计 [千克]；
                      eFault 为锁存回放；ePhaseBad 为非法相位兜底专用成员（R128）。
  修订记录 Revision  :
    2026-11-20  v1.0.0  R56 首版（批 4 · 序号 16）
    2026-11-21  v1.0.1  R57 返修：空闲相 / 失能迁移 / 故障锁存三路径输出安全侧归零
  ==================================================================
*)

TYPE E_DL_LwfPhase :
(
    eIdle   := 0,  // 空闲：等启动沿 / idle, waiting for the start edge
    eDose   := 10, // 给料：PI 闭环与批量累计 / dosing, the PI loop and the batch accumulation
    eRefill := 20, // 补料：计量冻结，等补料完成 / refilling, the metering freezes until the refill completes
    eDone   := 30, // 批次完成：驻留等复位或新启动 / done, held until reset or a new start
    eFault  := 90  // 故障：成因锁存 / fault, the cause is latched
);
END_TYPE

TYPE E_DL_LwfFault :
(
    eNone         := 0, // 无成因 / no cause
    eNoLossRate   := 1, // 输出非零而速率长期为零（故障级，与 bError 配对）/ a nonzero output with a void loss rate, fault grade paired with bError
    eWeightNoise  := 2, // 称重突跳超物理限（故障级，与 bError 配对）/ a weight jump beyond the physical limit, fault grade paired with bError
    eRefillTimeout:= 3, // 补料超时（故障级，与 bError 配对）/ the refill timed out, fault grade paired with bError
    eSensorBad    := 4, // 称重非有限或组态非法（故障级，与 bError 配对）/ the weight is non finite or the config illegal, fault grade paired with bError
    ePhaseBad     := 5  // 非法相位兜底（故障级，与 bError 配对）/ illegal phase fallback, fault grade paired with bError
);
END_TYPE

FUNCTION_BLOCK FB_DL_LossInWeightFeeder
VAR_INPUT
    bEnable     : BOOL := TRUE;    // 使能，失能时停给料回空闲 [-] / enable, the feeding stops when disabled
    bReset      : BOOL := FALSE;   // 复位上升沿清故障锁存与批量累计 [-] / reset rising edge clears the fault latch and the batch accumulation
    bStart      : BOOL := FALSE;   // 批次启动脉冲，上升沿受理 [-] / the batch start pulse, accepted on the rising edge
    bRefillDone : BOOL := FALSE;   // 补料完成脉冲（外部给出）[-] / the refill done pulse from the outside
    fWeightKg   : LREAL := 100.0;  // 称重实测 [千克] / the measured weight [kilogram]
    fRateSp     : LREAL := 10.0;   // 目标给料速率 [千克每小时]，域 大于零 / the target feed rate [kilogram per hour], domain above zero
    fKp         : LREAL := 2.0;    // PI 比例增益 [输出每速率误差] / the PI proportional gain [output per rate error]
    fTi         : LREAL := 30.0;   // PI 积分时间 [秒]，域 大于零 / the PI integral time [second], domain above zero
    fOutMax     : LREAL := 100.0;  // 输出上限 [百分比] / the output ceiling [percent]
    fRateFiltT  : LREAL := 2.0;    // 速率低通时间常数 [秒]，0 = 直通 / the rate low pass time constant [second], zero is a passthrough
    fNoiseLim   : LREAL := 500.0;  // 称重突跳物理限（速率口径）[千克每小时] / the weight jump physical limit in rate terms [kilogram per hour]
    fLowWeightKg: LREAL := 20.0;   // 低料位补料阈值 [千克] / the low weight refill threshold [kilogram]
    fBatchTarget: LREAL := 500.0;  // 批量目标 [千克]，域 大于零 / the batch target [kilogram], domain above zero
    tRefillTo   : TIME := T#120S;  // 补料超时窗 [毫秒]，域 大于 tNoRateTo / the refill timeout window, above the no rate window
    tNoRateTo   : TIME := T#10S;   // 无速率确认窗 [毫秒]，域 大于零 / the no rate confirm window [millisecond], domain above zero
    fDtS        : LREAL := 0.1;    // 调用周期 [秒]，域 大于零 / the call period [second], domain above zero
END_VAR
VAR_OUTPUT
    fRateOut  : LREAL := 0.0;  // 给料输出（PI 后，0..上限）[百分比] / the feed output after the PI [percent]
    bDosing   : BOOL := FALSE; // 给料中（相位派生电平）[-] / dosing, a phase derived level
    bRefilling: BOOL := FALSE; // 补料中（相位派生电平）[-] / refilling, a phase derived level
    fBatchAcc : LREAL := 0.0;  // 批量累计 [千克] / the batch accumulation [kilogram]
    ePhase    : E_DL_LwfPhase := E_DL_LwfPhase.eIdle; // 相位出口 [枚举] / phase outlet [enum]
    eFault    : E_DL_LwfFault := E_DL_LwfFault.eNone; // 成因出口，锁存回放 [枚举] / cause outlet replayed from the latch [enum]
    bError    : BOOL := FALSE; // 故障锁存标志 [-] / fault latch flag
END_VAR
VAR
    rtStart   : R_TRIG; // 启动沿检测，段 0 无条件刷新 / start edge, refreshed unconditionally in segment zero
    rtRefillD : R_TRIG; // 补料完成沿检测，段 0 无条件刷新 / refill done edge, refreshed unconditionally in segment zero
    rtReset   : R_TRIG; // 复位沿检测，段 0 无条件刷新 / reset edge, refreshed unconditionally in segment zero
    tonRefill : TON;    // 补料超时窗，段 0 无条件刷新 / the refill timeout window, refreshed unconditionally
    tonNoRate : TON;    // 无速率确认窗，段 0 无条件刷新 / the no rate confirm window, refreshed unconditionally
    _ePhase   : E_DL_LwfPhase := E_DL_LwfPhase.eIdle; // 内部相位，CASE 唯一写入目标 / internal phase, the only CASE write target
    _eFaulC   : E_DL_LwfFault := E_DL_LwfFault.eNone; // 故障级成因，锁存至复位沿 / fault cause, latched until the reset edge
    _bFault   : BOOL := FALSE; // 故障锁存位 [-] / fault latch bit
    _bInit    : BOOL := FALSE; // 首扫初始化完成标志（R310）/ first scan initialisation flag
    _bCfgOk   : BOOL := FALSE; // 组态参数域内 [-] / the configuration is inside the domain
    _bInOk    : BOOL := FALSE; // 称重有限 [-] / the weight is finite
    _fWPrev   : LREAL := 0.0;  // 上拍称重快照 [千克] / previous scan weight snapshot [kilogram]
    _fRateRaw : LREAL := 0.0;  // 原始失重速率 [千克每小时] / the raw loss rate [kilogram per hour]
    _fRateF   : LREAL := 0.0;  // 滤后失重速率 [千克每小时] / the filtered loss rate [kilogram per hour]
    _fE       : LREAL := 0.0;  // 速率误差 [千克每小时] / the rate error [kilogram per hour]
    _fI       : LREAL := 0.0;  // 积分项保持量 [百分比] / the integral term holder [percent]
    _fUPre    : LREAL := 0.0;  // 限幅前输出 [百分比] / the pre clamp output [percent]
    _fW       : LREAL := 0.0;  // 一阶低通权 [无量纲] / the first order weight
END_VAR

// 段 0｜定时器与沿检测无条件周期刷新（禁入分支），IN 只串相位闸与故障闸（FB50-1）/ segment 0, unconditional refresh, no instance call inside a branch
rtStart(CLK := bStart); // 启动沿 / the start edge
rtRefillD(CLK := bRefillDone); // 补料完成沿 / the refill done edge
rtReset(CLK := bReset); // 复位沿 / the reset edge
tonRefill(IN := (_ePhase = E_DL_LwfPhase.eRefill) AND (NOT _bFault), PT := tRefillTo); // 补料超时窗，IN 串补料相闸 / the refill timeout with the refill phase gate
tonNoRate(IN := (_ePhase = E_DL_LwfPhase.eDose) AND (fRateOut > 1.0) AND (NOT _bFault), PT := tNoRateTo); // 无速率确认窗，IN 串给料相闸与输出非零判据 / the no rate window with the dose phase gate

// 段 1｜首扫初始化（R310）/ segment 1, first scan initialisation
IF NOT _bInit THEN // 首扫一拍 / the very first scan
    _bInit := TRUE; // 置首扫完成标志 / raise the first scan flag
    _ePhase := E_DL_LwfPhase.eIdle; // 相位从空闲起步 / the phase starts from idle
    _eFaulC := E_DL_LwfFault.eNone; // 故障级成因清零 / clear the fault cause
    _bFault := FALSE; // 故障锁存清零 / clear the fault latch
    _fWPrev := fWeightKg; // 快照取当拍 / the snapshot takes this scan
END_IF

// 段 2｜复位沿作用域：清锁存 / 迁相位 / 清批量累计与积分（三项逐项声明）/ segment 2, reset edge scope declared item by item
IF rtReset.Q THEN // 复位沿 / the reset edge
    _bFault := FALSE; // 作用域一：清故障锁存 / scope one, clear the fault latch
    _eFaulC := E_DL_LwfFault.eNone; // 作用域一：清故障级成因 / scope one, clear the fault cause
    _ePhase := E_DL_LwfPhase.eIdle; // 作用域二：迁回空闲相 / scope two, migrate back to idle
    fBatchAcc := 0.0; // 作用域三：清批量累计 / scope three, clear the batch accumulation
    _fI := 0.0; // 作用域三：清积分项 / scope three, clear the integral term
    _fRateF := 0.0; // 作用域三：清滤后速率 / scope three, clear the filtered rate
END_IF

// 段 3｜组态与输入域闸（R151 全覆盖）/ segment 3, the configuration and input domain gates
_bInOk := (fWeightKg = fWeightKg) AND ((fWeightKg - fWeightKg) = (fWeightKg - fWeightKg)); // 称重有限性 / the weight finiteness
_bCfgOk := (fRateSp > 0.0) AND (fRateSp = fRateSp) AND (fKp > 0.0) AND (fKp = fKp) AND (fTi > 0.0) AND (fTi = fTi) AND (fOutMax > 0.0) AND (fOutMax = fOutMax) AND (fRateFiltT >= 0.0) AND (fRateFiltT = fRateFiltT) AND (fNoiseLim > 0.0) AND (fNoiseLim = fNoiseLim) AND (fBatchTarget > 0.0) AND (fBatchTarget = fBatchTarget) AND (tRefillTo > T#0S) AND (tNoRateTo > T#0S) AND (tRefillTo > tNoRateTo) AND (fDtS > 0.0) AND (fDtS = fDtS); // 组态参数域判定（含 R100 配比）/ the configuration verdict with the window pairing
IF (NOT _bInOk) OR (NOT _bCfgOk) THEN // 输入非有限或组态非法 / a non finite input or an illegal configuration
    IF NOT _bFault THEN // 未锁存才迁移（防同拍抹除）/ migrate only while unlatched
        _bFault := TRUE; // 置故障锁存 / raise the fault latch
        _eFaulC := E_DL_LwfFault.eSensorBad; // 故障级成因（R45 配对 bError）/ the fault cause paired with bError
        _ePhase := E_DL_LwfPhase.eFault; // 迁故障相 / migrate to the fault phase
    END_IF
END_IF

// 段 4｜失重速率计算（含噪声闸）：快照推进无条件执行，防恢复时速率踢 / segment 4, the loss rate computation with the noise gate, the snapshot advances unconditionally
_fRateRaw := 0.0; // 原始速率预置零 / preset the raw rate to zero
IF _bInOk AND _bCfgOk THEN // 输入与组态合法 / the input and the config are legal
    _fRateRaw := (_fWPrev - fWeightKg) / fDtS * 3600.0; // 失重速率 = 负变化 / 周期，转千克每小时（除子为周期已证大于零）/ the loss rate converted to kilogram per hour with a proven divisor
    IF ABS(_fRateRaw) > fNoiseLim THEN // 称重突跳超物理限 / the weight jump exceeds the physical limit
        IF NOT _bFault THEN // 未锁存才迁移 / migrate only while unlatched
            _bFault := TRUE; // 置故障锁存 / raise the fault latch
            _eFaulC := E_DL_LwfFault.eWeightNoise; // 故障级成因（R45 配对 bError）/ the fault cause paired with bError
            _ePhase := E_DL_LwfPhase.eFault; // 迁故障相 / migrate to the fault phase
        END_IF
        _fRateRaw := 0.0; // 本拍噪声样本不参与 / the noisy sample does not participate
    END_IF
END_IF
_fWPrev := fWeightKg; // 快照推进（无条件）/ the snapshot advances unconditionally

// 段 5｜相位机：ENUM + CASE，含 ELSE 非法相位兜底（R128）/ segment 5, the phase machine with an ELSE fallback
CASE _ePhase OF
E_DL_LwfPhase.eIdle: // 空闲相：等启动沿 / the idle phase, waiting for the start edge
    fRateOut := 0.0; // 空闲相输出强制安全侧归零（v1.0.1 返修）/ the outlet is force-zeroed on the safe side while idle (v1.0.1 fix)
    IF bEnable AND (NOT _bFault) AND rtStart.Q THEN // 启动沿受理 / the start edge is accepted
        _ePhase := E_DL_LwfPhase.eDose; // 迁给料相 / migrate to the dose phase
    END_IF

E_DL_LwfPhase.eDose: // 给料相：PI 闭环 + 批量累计 + 低料位切换 / the dose phase, the PI loop, the accumulation and the refill switch
    IF NOT bEnable THEN // 失能 / disabled
        fRateOut := 0.0; // 迁移前先归零（安全侧，v1.0.1 返修）/ zeroed on the safe side before the migration (v1.0.1 fix)
        _ePhase := E_DL_LwfPhase.eIdle; // 回空闲相 / back to idle
    ELSE // 正常给料 / the normal feeding
        IF fRateFiltT > 0.0 THEN // 低通开启 / the low pass is on
            _fW := fDtS / (fDtS + fRateFiltT); // 一阶低通权，除子已证大于零 / the first order weight with a proven divisor
            _fRateF := _fRateF + _fW * (_fRateRaw - _fRateF); // 速率低通推进 / advance the rate low pass
        ELSE // 直通口径 / the passthrough
            _fRateF := _fRateRaw; // 原始速率直通 / the raw rate passes through
        END_IF
        fBatchAcc := fBatchAcc + _fRateF * fDtS / 3600.0; // 批量累计（千克每小时 × 秒 / 3600）/ accumulate the batch
        _fE := fRateSp - _fRateF; // 速率误差 / the rate error
        _fUPre := fKp * _fE + _fI; // 限幅前输出（比例 + 积分保持量）/ the pre clamp output
        IF NOT ((_fUPre >= fOutMax) AND (_fE > 0.0)) THEN // 未沿误差方向饱和才积分（抗 windup）/ the integration is gated against the saturation direction
            _fI := _fI + (fKp / fTi) * _fE * fDtS; // 积分推进，除子为积分时间已证大于零 / the integral step with the proven divisor
        END_IF
        _fUPre := fKp * _fE + _fI; // 积分后重算 / recompute after the integral
        IF _fUPre < 0.0 THEN // 下限钳零 / clamp the floor to zero
            fRateOut := 0.0; // 输出归零 / the output is zeroed
        ELSIF _fUPre > fOutMax THEN // 上限钳制 / clamp the ceiling
            fRateOut := fOutMax; // 钳到上限 / clamp to the ceiling
        ELSE // 域内 / inside the domain
            fRateOut := _fUPre; // 直接出口 / straight to the outlet
        END_IF
        IF fBatchAcc >= fBatchTarget THEN // 批量达标 / the batch target is reached
            _ePhase := E_DL_LwfPhase.eDone; // 迁完成相 / migrate to the done phase
        ELSIF fWeightKg <= fLowWeightKg THEN // 低料位触发补料 / the low weight triggers the refill
            fRateOut := 0.0; // 补料前输出归零（冻结语义）/ the output zeroes before the refill
            _ePhase := E_DL_LwfPhase.eRefill; // 迁补料相 / migrate to the refill phase
        ELSIF tonNoRate.Q THEN // 输出非零而速率长期为零 / a nonzero output with a void rate
            _bFault := TRUE; // 置故障锁存 / raise the fault latch
            _eFaulC := E_DL_LwfFault.eNoLossRate; // 故障级成因（R45 配对 bError）/ the fault cause paired with bError
            _ePhase := E_DL_LwfPhase.eFault; // 迁故障相 / migrate to the fault phase
        END_IF
    END_IF

E_DL_LwfPhase.eRefill: // 补料相：计量冻结，等完成沿（退出条件 ≥2：完成沿 / 超时 / 失能，R98）/ the refill phase with the metering frozen, at least two exit conditions
    fRateOut := 0.0; // 输出保持归零（R191 冻结语义显式声明）/ the output holds zeroed per the declared frozen semantics
    bRefilling := TRUE; // 补料指示 / the refilling indicator
    IF NOT bEnable THEN // 失能 / disabled
        _ePhase := E_DL_LwfPhase.eIdle; // 回空闲相 / back to idle
    ELSIF rtRefillD.Q THEN // 补料完成沿 / the refill done edge
        _fI := 0.0; // 积分项清零（恢复后重新爬坡）/ clear the integral for a fresh ramp
        _ePhase := E_DL_LwfPhase.eDose; // 迁回给料相 / migrate back to the dose phase
    ELSIF tonRefill.Q THEN // 补料超时 / the refill timed out
        _bFault := TRUE; // 置故障锁存 / raise the fault latch
        _eFaulC := E_DL_LwfFault.eRefillTimeout; // 故障级成因（R45 配对 bError）/ the fault cause paired with bError
        _ePhase := E_DL_LwfPhase.eFault; // 迁故障相 / migrate to the fault phase
    END_IF

E_DL_LwfPhase.eDone: // 完成相：输出归零，等复位或新启动 / the done phase, the output zeroes until reset or a new start
    fRateOut := 0.0; // 输出归零 / the output is zeroed
    IF NOT bEnable THEN // 失能 / disabled
        _ePhase := E_DL_LwfPhase.eIdle; // 回空闲相 / back to idle
    ELSIF rtStart.Q THEN // 新启动沿 / a new start edge
        fBatchAcc := 0.0; // 批量累计清零 / clear the batch accumulation
        _fI := 0.0; // 积分项清零 / clear the integral term
        _ePhase := E_DL_LwfPhase.eDose; // 迁给料相 / migrate to the dose phase
    END_IF

E_DL_LwfPhase.eFault: // 故障相：输出归零，成因锁存，等复位沿 / the fault phase, the output zeroes until the reset edge
    fRateOut := 0.0; // 输出安全侧归零 / the output takes the safe side zero
    IF NOT bEnable THEN // 失能 / disabled
        _ePhase := E_DL_LwfPhase.eIdle; // 迁未使能相 / migrate to idle
    END_IF

ELSE // 非法相位兜底（R128）/ the illegal phase fallback
    _bFault := TRUE; // 置故障锁存 / raise the fault latch
    _eFaulC := E_DL_LwfFault.ePhaseBad; // 故障级成因（R45 配对 bError）/ the fault cause paired with bError
    _ePhase := E_DL_LwfPhase.eFault; // 迁故障相 / migrate to the fault phase
END_CASE

// 段 6｜统一出口 / segment 6, the unified outlet
IF _bFault THEN // 故障锁存优先 / the fault latch takes priority
    fRateOut := 0.0; // 故障拍输出安全侧归零（v1.0.1 返修）/ the outlet is zeroed on the safe side while faulted (v1.0.1 fix)
    eFault := _eFaulC; // 故障级成因锁存回放（R152）/ the fault cause replayed from the latch
ELSE
    eFault := E_DL_LwfFault.eNone; // 无锁存即无成因 / no latch, no cause
END_IF
bDosing := (_ePhase = E_DL_LwfPhase.eDose); // 给料指示（相位派生）/ the dosing indicator derived from the phase
bRefilling := (_ePhase = E_DL_LwfPhase.eRefill); // 补料指示（相位派生）/ the refilling indicator derived from the phase
ePhase := _ePhase; // 相位出口单点映射 / single point phase outlet mapping
bError := _bFault; // 故障标志与锁存位同源 / the fault flag shares the latch source
END_FUNCTION_BLOCK

(* ---- FB_DL_LowPassFilter.st ---- *)
(*==============================================================================
 * 组件名称 (Component)  : FB_DL_LowPassFilter
 * 所属子库 (Sublibrary) : DL_Algo
 * 当前版本 (Version)    : 1.0.0
 * 兼容性   (Platform)   : CODESYS 3.5 / TwinCAT 3 / 汇川 InoProShop / Machine Expert
 *                         仅依赖 Standard.library（MIN / MAX / ABS），零厂商方言
 * 功能描述 (Function)   : 一阶惯性低通数字滤波器（PT1 / LGF PT1 语义）。
 *                         递推式 fOut := fOut + fAlpha*(fIn - fOut)，
 *                         其中 fAlpha := fDt / (fTf + fDt)；时间常数 tTimeConst
 *                         运行中可调，变更即时重算 fAlpha；tTimeConst = 0 直通；
 *                         首扫与 bTrack 跟踪均无滞后，投切无扰动。
 *                         现场用途：温度 / 压力 / 流量模拟量采集降噪。
 * 开源溯源 (Origin)     : 原创实现。算法思想源自 LGF PT1 与模板库
 *                         05-algorithm-templates.md 的 FB_LowPassFilter 结构，
 *                         按本库故障码体系（16#0002_xxxx）重写并加严。
 * 设计验证 (Verified)   : fT1=0.1s、fDt=0.01s、阶跃 0->1（python 6 位小数）：
 *                         fAlpha=0.090909；第 1 拍 fOut=0.090909；
 *                         第 10 拍 fOut=0.614457；第 50 拍 fOut=0.991481。
 * 验收向量 (Acceptance) :
 *   V1 fT1=0.1s fDt=0.01s 输入恒 1.0：第 1 拍 fOut≈0.090909（容差 1E-4）
 *   V2 同 V1：第 10 拍 fOut≈0.614457（容差 1E-4）
 *   V3 同 V1：第 50 拍 fOut≈0.991481（容差 1E-4）
 *   V4 tTimeConst=T#0S：任意输入当拍直通，fOut=fIn、fAlpha=1.0
 *   V5 bTrack=TRUE fTrackValue=42.0：当拍 fOut=42.0 且无爬升过程
 *   V6 fIn 非有限值：本拍拒绝更新保持上拍输出，uErrorId=16#0002_0004
 * 本文件内含       : TYPE  E_DL_LpfState（配套枚举，归属 DL_Algo）
 *                    FB    FB_DL_LowPassFilter
 * 依赖     (Depends)    : 无 DL_ 内部依赖；Standard.library 数学算符
 * 红线自检 (Redline)    : R1 ✓ 零全局变量表与外部变量引用 ｜ R2 ✓ 零物理 IO 地址直写
 *                         R3 ✓ 纯 IEC 61131-3 ｜ R4 ✓ 钳位+容差+非有限值拒绝+防除零
 *                         R5 ✓ 全变量中英双语同行注释 ｜ R6 ✓ 四态 ENUM+CASE+ELSE
 *                         R7 N/A（无定时器与边沿检测实例）
 * 修订历史 (Revision)   :
 *   2026-11-15  v1.0.0  首版入库（Round 04 · Phase 3 · DL_Algo 批次）
 *============================================================================*)

(*-----------------------------------------------------------------------------
 * 调用示例 (Instance guide)：
 *   声明于调用方 FB 的 VAR 区：fbLpf : FB_DL_LowPassFilter;
 *   每周期调用：fbLpf(bEnable := TRUE, fIn := stPv.fRaw,
 *                     tTimeConst := T#1S, tSampleTime := T#100MS);
 *   取用输出：  stPv.fFiltered := fbLpf.fOut;
 * 现场调参指引：温度回路 tTimeConst 取 1 到 3 秒，压力回路取 0.3 到 1 秒；
 *   投入调节回路前先用 bTrack 跟踪当前过程值，切换瞬间输出无跳变。
 *----------------------------------------------------------------------------*)

(*-----------------------------------------------------------------------------
 * 枚举: E_DL_LpfState（归属 DL_Algo，与 FB_DL_LowPassFilter 同文件）
 * 含义: 低通滤波状态机离散状态。纯线性滤波采用「状态派生 + CASE 覆盖 + ELSE」
 *       结构：状态由使能 / 跟踪 / 首扫信号派生，CASE 保证每态行为显式可审计。
 *----------------------------------------------------------------------------*)
TYPE E_DL_LpfState :
(
    eInit  := 0,    // 首扫态：输出直接采样输入，bValid=FALSE，无历史瞬态 / First scan: output tracks input directly, bValid=FALSE
    eRun   := 10,   // 运行态：按 fAlpha 递推滤波，参数变更即时生效 / Running: recursive filtering with live fAlpha, parameter changes apply at once
    eTrack := 20,   // 跟踪态：输出立即跟随 fTrackValue，内部历史同步 / Tracking: output follows fTrackValue instantly, states synchronized
    eFault := 99    // 故障兜底态：非法状态进入，输出安全值并置故障码 / Fault fallback: entered from illegal states, safe output plus error code
);
END_TYPE

(*==============================================================================
 * 功能块: FB_DL_LowPassFilter
 * 调用约定: 每个采样周期无条件调用一次；tSampleTime 由调用方显式给定，
 *           严禁依赖隐式扫描周期做滤波递推；多实例可并行互不干扰。
 * 滞后披露: 输出对阶跃的 63.2% 响应时间约等于 tTimeConst（离散近似），
 *           tTimeConst 越大越平滑、相位滞后越大，选型需与采样周期匹配。
 *============================================================================*)
FUNCTION_BLOCK FB_DL_LowPassFilter
VAR_INPUT
    bEnable     : BOOL := FALSE;      // 使能，FALSE 时输出直通原始输入 / Enable, FALSE passes raw input straight through
    fIn         : REAL := 0.0;        // 原始采样输入 [EU] / Raw sampling input [EU]
    tTimeConst  : TIME := T#1S;       // 滤波时间常数 [s]，T#0S = 直通 / Filter time constant [s], T#0S = pass-through
    tSampleTime : TIME := T#100MS;    // 采样周期 [s 口径换算]，小于 10ms 钳位 / Sampling period, clamped to 10ms minimum
    bTrack      : BOOL := FALSE;      // 跟踪使能，TRUE 时输出立即跟随跟踪值 / Track enable, TRUE makes output follow track value instantly
    fTrackValue : REAL := 0.0;        // 跟踪目标值 [EU]，无扰投切用 / Track target value [EU], for bumpless transfer
END_VAR
VAR_OUTPUT
    fOut        : REAL;               // 滤波输出 [EU] / Filtered output [EU]
    fAlpha      : REAL;               // 当前滤波系数 [0..1]，诊断用 / Current filter coefficient [0..1], diagnostic
    bValid      : BOOL;               // 输出有效标志，首扫未完成时为 FALSE / Output valid flag, FALSE before first scan completes
    bError      : BOOL;               // 故障标志，与 uErrorId 联动 / Fault flag, coupled with uErrorId
    uErrorId    : UDINT;              // 故障码，0 = 无故障 / Error code, 0 = no error
END_VAR
VAR
    fTfEff      : REAL;               // 钳位后的生效时间常数 [s] / Effective clamped time constant [s]
    fDt         : REAL;               // 采样周期秒值 [s] / Sampling period in seconds [s]
    fTfRaw      : REAL;               // 时间常数换算秒值（钳位前）[s] / Time constant in seconds before clamping [s]
    eState      : E_DL_LpfState;      // 状态机当前状态 / Current state of the state machine
END_VAR
VAR CONSTANT
    DL_LPF_TF_MAX  : REAL := 3600.0;  // 时间常数上限 [s]，超限钳位防极端迟滞 / Time constant upper clamp [s], prevents extreme lag
    DL_LPF_DT_MIN  : REAL := 0.01;    // 采样周期防御下限 [s] / Defensive sampling period lower bound [s]
    DL_LPF_INF_MAX : REAL := 1.0E30;  // 有限值判定幅值上限 [EU] / Magnitude bound for finite-value check [EU]
END_VAR

(*------------------------------------------------------------------------------
 * 段 1｜参数钳位（不中断扫描）：采样周期下限与时间常数越界只置码修正
 *      Parameter clamping without scan interruption: period floor and constant range
 *-----------------------------------------------------------------------------*)
uErrorId := 16#0002_0000;

IF tSampleTime < T#10MS THEN
    fDt      := DL_LPF_DT_MIN;                       // 周期过小钳位到 10ms / Too small period clamped to 10ms
    uErrorId := 16#0002_0002;                        // 采样周期非法已钳位 / Invalid sampling period clamped
ELSE
    fDt := TIME_TO_REAL(tSampleTime) / 1000.0;       // TIME 换算秒值 / Convert TIME to seconds
END_IF

fTfRaw := TIME_TO_REAL(tTimeConst) / 1000.0;         // 时间常数换算秒值 / Convert time constant to seconds

IF (fTfRaw < 0.0) OR (fTfRaw > DL_LPF_TF_MAX) THEN
    fTfEff   := MIN(MAX(fTfRaw, 0.0), DL_LPF_TF_MAX); // 双侧钳位到合法域 / Two-sided clamp into valid range
    uErrorId := 16#0002_1001;                        // 时间常数非法已钳位 / Invalid time constant clamped
ELSE
    fTfEff := fTfRaw;                                // 合法参数原值生效 / Valid parameter applied as-is
END_IF

(*------------------------------------------------------------------------------
 * 段 2｜滤波系数计算（防除零 + 显式区间约束）：fAlpha = fDt/(fTf+fDt)
 *      Filter coefficient with divide-by-zero guard and explicit interval
 *      tTimeConst=0 时 fAlpha=1.0，天然直通，与 V4 向量对应
 *-----------------------------------------------------------------------------*)
IF fTfEff <= 1.0E-6 THEN
    fAlpha := 1.0;                                   // 零时间常数直通系数 / Pass-through coefficient for zero constant
ELSE
    fAlpha := MIN(MAX(fDt / (fTfEff + fDt), 0.0), 1.0); // 系数显式约束在 0 与 1 之间 / Coefficient constrained into 0..1
END_IF

(*------------------------------------------------------------------------------
 * 段 3｜非有限值防御：拒绝本拍更新、保持上一拍输出（公共故障码）
 *      Non-finite defense: reject this cycle, hold previous output
 *-----------------------------------------------------------------------------*)
IF (fIn <> fIn) OR (ABS(fIn) > DL_LPF_INF_MAX) THEN
    uErrorId := 16#0002_0004;                        // 输入非有限值已拒绝 / Non-finite input rejected
    bValid   := FALSE;
    bError   := TRUE;
    RETURN;
END_IF

(*------------------------------------------------------------------------------
 * 段 4｜主状态机（红线 R6）：状态派生 + CASE 覆盖 + ELSE 兜底
 *      Main state machine: state derived from signals, CASE covered with ELSE
 *-----------------------------------------------------------------------------*)
IF bTrack THEN
    eState := eTrack;                                // 跟踪请求优先级最高 / Track request has highest priority
ELSIF eState = eInit THEN
    eState := eInit;                                 // 首扫态保持，不被运行派生覆盖 / First scan state preserved from override
ELSIF eState = eFault THEN
    IF NOT bEnable THEN
        eState := eInit;                             // 使能跌落提供故障恢复路径 / Disabled input provides fault recovery path
    ELSE
        eState := eFault;                            // 故障态保持直至调用方处置 / Fault state holds until caller intervenes
    END_IF
ELSE
    eState := eRun;                                  // 常规运行态派生 / Normal running state derived
END_IF

CASE eState OF

    eInit:
        (* 首扫直接采样：输出等于输入，无历史瞬态（与验收 V5 等价的天然行为） *)
        (* First scan samples directly: output equals input, no historical transient *)
        fOut   := fIn;
        bValid := FALSE;                             // 首扫未完成，输出尚不可信 / First scan unfinished, output not trustworthy yet
        eState := eRun;                              // 下一拍进入运行态 / Move to running state next cycle

    eTrack:
        (* 无扰跟踪：输出立即跟随跟踪值，滤波历史同步置位，回自动无跳变 *)
        (* Bumpless tracking: output follows track value, filter state synchronized *)
        fOut   := fTrackValue;
        bValid := TRUE;
        eState := eRun;

    eRun:
        IF NOT bEnable THEN
            (* 使能失效语义：直通原始输入，系数保持显示但不参与递推 *)
            (* Disabled semantics: pass raw input through, coefficient kept for display only *)
            fOut   := fIn;
            bValid := FALSE;
        ELSE
            (* 一阶低通递推：fOut += (fIn - fOut) * fAlpha，fAlpha 已在段 2 确定 *)
            (* First-order recursion: fOut += (fIn - fOut) * fAlpha *)
            fOut   := fOut + (fIn - fOut) * fAlpha;
            bValid := TRUE;
        END_IF

    eFault:
        (* 故障兜底：输出保持安全值 0，等待调用方修正参数后重新派生 *)
        (* Fault fallback: output holds safe value 0 until caller fixes parameters *)
        fOut   := 0.0;
        bValid := FALSE;

    ELSE
        (* 非法状态拦截：任何未定义枚举值一律进故障态并置公共兜底码 *)
        (* Illegal state interception: undefined enum values go to fault with code *)
        eState   := eFault;
        fOut     := 0.0;
        bValid   := FALSE;
        uErrorId := 16#0002_0005;

END_CASE;

(* 故障标志统一出口：与故障码严格联动，0 即无故障 *)
(* Unified fault flag outlet: strictly coupled with error code, zero means healthy *)
bError := (uErrorId <> 16#0002_0000);
END_FUNCTION_BLOCK

(* ---- FB_DL_MracAdaptiveCtrl.st ---- *)
(*
  ==================================================================
  组件名 Component  : FB_DL_MracAdaptiveCtrl
  分类   Category   : DL_Algo
  复杂度 Complexity  : 重
  版本   Version    : 1.0.0
  功能   Purpose    : 模型参考自适应控制器（MRAC）。一阶参考模型
                      dModel/dt = (fRefCmd − Model)/Tm；跟踪误差 e = Model −
                      YMeas 驱动可调增益 σ 修正更新：dKp/dt = γ·e·fRefCmd −
                      σ·Kp（防参数漂移），增益钳位 [fKmin, fKmax]；控制输出
                      fU = Kp·fRefCmd。欧拉离散，步长 fDtSec 由调用方给定。
                      与 FB_DL_RlsEstimator 参数辨识分工互引。
  来源   Source     : self（MRAC 公开控制理论）
  溯源   Origin     : MIT 规则 MRAC 与 σ 修正为公开控制理论语义，clean-room
                      自研实现，未复制任何厂商私有库源码。
  平台   Platform   : 纯 IEC 61131-3，CODESYS / TwinCAT / InoProShop 通用
  分工声明 Split     : 与 FB_DL_RlsEstimator 分工——后者做递推参数辨识，
                      本件做参考模型驱动的在线增益自适应。
  作者   Author     : 道莅代码库 · PLC 编程专家（R59）
  ------------------------------------------------------------------
  边界 Boundary     :
                      一 非有限/组态闸（自反双判据 + 域闸）：fDtSec ∉ (0,0.1]
                         或 Tm ≤ eps 或入参非有限 → bBad 置位（本库纪律②），
                         状态冻结、fU 安全侧零；
                      二 增益硬钳位 [fKmin, fKmax] 单点回夹（防自适应发散）；
                      三 复位沿：Model/Kp/输出全清（解除路径 = bReset 沿，
                         R188）；
                      四 首拍初始化（R310 真实使用）：Model 预置取当前测量
                         值（状态从测量起跳，防首拍误差尖峰）；
                      五 无全局变量、无外部变量声明、无物理地址寻址。
  修订记录 Revision  :
    2026-11-21  v1.0.0  R59 首版（批 3 · 序号 11）
  ==================================================================
*)

FUNCTION_BLOCK FB_DL_MracAdaptiveCtrl
VAR_INPUT
    fRefCmd : LREAL := 0.0;  // 参考指令 [工程单位] / the reference command [engineering unit]
    fYMeas  : LREAL := 0.0;  // 被控量测量 [工程单位] / the plant measurement [engineering unit]
    fDtSec  : LREAL := 0.01; // 离散步长 [秒]，域 (0, 0.1] / the discrete step [second]
    fTmSec  : LREAL := 0.5;  // 参考模型时间常数 [秒]，域 > eps / the model time constant [second]
    fGamma  : LREAL := 0.5;  // 自适应增益 [1/(单位·秒)] / the adaptive gain
    fSigma  : LREAL := 0.01; // σ 修正系数 [1/秒]，防漂移 / the sigma modification, anti drift
    fKmin   : LREAL := -10.0; // 增益下钳位 [无量纲] / the gain clamp floor
    fKmax   : LREAL := 10.0;  // 增益上钳位 [无量纲] / the gain clamp ceiling
    bEnable : BOOL := FALSE;  // 使能，失能状态冻结输出零 [-] / the enable, disabling freezes and zeroes
    bReset  : BOOL := FALSE;  // 复位上升沿清状态 [-] / the reset rising edge clears the states
END_VAR
VAR_OUTPUT
    fU      : LREAL := 0.0; // 控制输出 [工程单位] / the control outlet [engineering unit]
    fModelY : LREAL := 0.0; // 参考模型输出 [工程单位] / the model outlet [engineering unit]
    fETrack : LREAL := 0.0; // 跟踪误差（Model − YMeas）[工程单位] / the tracking error [engineering unit]
    fKp     : LREAL := 0.0; // 可调增益实时值 [无量纲] / the adaptive gain live value
    bBad    : BOOL := FALSE; // 非有限/组态闸实时标志 [-] / the non finite or config gate flag
    bValid  : BOOL := FALSE; // 输出可用标志 [-] / the output usable flag
END_VAR
VAR CONSTANT
    DL_MRA_EPS   : LREAL := 1.0E-9;  // 时间常数下阈值 [秒] / the time constant threshold
    DL_MRA_DTMAX : LREAL := 0.1;     // 步长上界 [秒] / the step ceiling
    DL_MRA_EMAX  : LREAL := 1.0E6;   // 跟踪误差钳位（数值防溢出）[工程单位] / the tracking error clamp, numeric
    DL_MRA_KMAXABS : LREAL := 1.0E6; // 自适应增益上界绝对值（R59 补：防 +Inf 穿闸）[—] / the absolute bound on the adaptive gain
END_VAR
VAR
    _fModel : LREAL := 0.0; // 参考模型状态 [工程单位] / the reference model state
    _fKp    : LREAL := 0.0; // 可调增益状态 [无量纲] / the adaptive gain state
    _fE     : LREAL;        // 跟踪误差工作量（含钳位）[工程单位] / the tracking error work value, clamped
    _bFin   : BOOL;         // 入参有限工作量 [-] / the input finiteness work flag
    _bCfg   : BOOL;         // 组态域工作量 [-] / the config domain work flag
    _bInit  : BOOL := FALSE; // 首拍初始化标志（R310，真实使用：模型起跳测量值）/ the first scan flag, real use
    rtReset : R_TRIG;        // 复位沿，段 0 无条件刷新 / the reset edge
END_VAR

// 段 0｜沿检测无条件周期刷新（禁入分支，R7）/ segment 0, the unconditional refresh
rtReset(CLK := bReset); // 复位沿 / the reset edge

// 段 1｜复位沿作用域：全状态清（解除路径 = bReset 沿，R188）/ segment 1, the reset edge scope
IF rtReset.Q THEN // 复位沿 / the reset edge
    _fModel := 0.0; // 模型状态清 / clear the model state
    _fKp := 0.0; // 增益状态清 / clear the gain state
    fModelY := 0.0; // 模型输出清 / clear the model outlet
    fKp := 0.0; // 增益出口清 / clear the gain outlet
    fU := 0.0; // 控制输出清（安全侧）/ clear the control, the safe side
    bValid := FALSE; // 有效降假 / drop the valid
END_IF

// 段 2｜首拍初始化（R310 真实使用路径）：模型起跳当前测量值 / segment 2, the first scan init, the model jump to the measurement
IF NOT _bInit THEN // 首拍一拍 / the first scan
    _bInit := TRUE; // 置首拍标志 / raise the flag
    _fModel := fYMeas; // 模型从测量起跳（防首拍误差尖峰）/ the model starts at the measurement
END_IF

// 段 3｜非有限与组态闸（边界一，实时标志非锁存）/ segment 3, the non finite and the config gate
_bFin := (fRefCmd = fRefCmd) AND ((fRefCmd - fRefCmd) = (fRefCmd - fRefCmd)) // 指令有限 / the command finite
    AND (fYMeas = fYMeas) AND ((fYMeas - fYMeas) = (fYMeas - fYMeas)) // 测量有限 / the measurement finite
    AND (fGamma = fGamma) AND ((fGamma - fGamma) = (fGamma - fGamma)) // 自适应增益有限 / the gain finite
    AND (fSigma = fSigma) AND ((fSigma - fSigma) = (fSigma - fSigma)) // σ 系数有限 / the sigma finite
    AND (fDtSec = fDtSec) AND ((fDtSec - fDtSec) = (fDtSec - fDtSec)) // 步长有限（R59 补）/ the step finite
    AND (fTmSec = fTmSec) AND ((fTmSec - fTmSec) = (fTmSec - fTmSec)) // 时间常数有限（R59 补）/ the time constant finite
    AND (fKmin = fKmin) AND (fKmax = fKmax) // 增益上下界有限（R59 补，防 +Inf 穿闸）/ the gain bounds finite
    AND (fKmin - fKmin = 0.0) AND (fKmax - fKmax = 0.0); // 界非无穷（R59 补）/ the bounds not infinite
_bCfg := (fDtSec > 0.0) AND (fDtSec <= DL_MRA_DTMAX) AND (fTmSec > DL_MRA_EPS) // 步长与时间常数域 / the step and the time constant domain
    AND (fKmin < fKmax) // 钳位序合理 / the clamp order sane
    AND (fKmax <= DL_MRA_KMAXABS); // 增益上界绝对值闸（R59 补）/ the absolute gain ceiling
bBad := (NOT _bFin) OR (NOT _bCfg); // 闸实时标志（R191 名实双出口）/ the gate flag

// 段 4｜自适应核心（使能且闸通过才推进；失能或闸拦状态冻结，边界一二）/ segment 4, the adaptive core
IF bEnable AND (NOT bBad) THEN // 有效推进窗 / the valid advance window
    _fModel := _fModel + (fDtSec * (fRefCmd - _fModel) / fTmSec); // 参考模型欧拉一步（除子 Tm 已闸）/ the model Euler step, divided by the gated Tm
    fModelY := _fModel; // 模型出口 / the model outlet
    _fE := _fModel - fYMeas; // 跟踪误差 / the tracking error
    IF _fE > DL_MRA_EMAX THEN // 误差上钳（数值防溢出）/ clamp the error up
        _fE := DL_MRA_EMAX; // 夹到上界 / clamp to the ceiling
    ELSIF _fE < -DL_MRA_EMAX THEN // 误差下钳 / clamp the error down
        _fE := -DL_MRA_EMAX; // 夹到下界 / clamp to the floor
    END_IF
    fETrack := _fE; // 误差出口（钳后口径）/ the error outlet, the clamped value
    _fKp := _fKp + (fDtSec * ((fGamma * _fE * fRefCmd) - (fSigma * _fKp))); // σ 修正增益更新 / the sigma modified gain update
    IF _fKp > fKmax THEN // 增益上钳（单点回夹）/ clamp the gain up
        _fKp := fKmax; // 夹到上界 / clamp to the ceiling
    ELSIF _fKp < fKmin THEN // 增益下钳 / clamp the gain down
        _fKp := fKmin; // 夹到下界 / clamp to the floor
    END_IF
    fKp := _fKp; // 增益出口 / the gain outlet
    fU := _fKp * fRefCmd; // 控制输出 / the control outlet
    bValid := TRUE; // 输出可用 / the output usable
ELSE // 失能或闸拦：输出安全侧零，状态冻结（边界一）/ disabled or gated, the safe zero and the frozen states
    fU := 0.0; // 控制输出安全零 / the safe zero
    fModelY := _fModel; // 模型出口保持冻结值 / the frozen model outlet
    fKp := _fKp; // 增益出口保持冻结值 / the frozen gain outlet
    fETrack := _fModel - fYMeas; // 误差出口保持观测（不推进）/ the observed error, not advanced
    IF NOT ((fETrack = fETrack) AND ((fETrack - fETrack) = (fETrack - fETrack))) THEN // 冻结出口非有限防护（R59 补）/ the frozen outlet finite guard
        fETrack := 0.0; // 非有限落安全零，不静默穿透 / non finite to the safe zero
    END_IF
    bValid := FALSE; // 可用降假 / drop the valid
END_IF
END_FUNCTION_BLOCK

(* ---- FB_DL_NotchFilter.st ---- *)
(*
    FB_DL_NotchFilter —— 二阶陷波滤波（中心频率与 Q 可调）
    ------------------------------------------------------------------
    分类      : DL_Algo / Filter
    前缀      : FB_DL_
    版本      : 1.0.0
    溯源      : T2-1 LGF · Measurement（只借「滤波归测量组」的分类事实）；
                陷波器双线性变换为公开数字信号处理公式，系数式、闸门顺序、码位分级
                100% 自有；clean-room 重写，未复制任何闭源厂商源码，
                参考实现仅限 MIT/Apache 许可
    平台      : 纯 IEC 61131-3，CODESYS V3.5+ / TwinCAT 3 / InoProShop 通用
    作者      : 道莅代码库 · PLC编程专家（R18）
    ------------------------------------------------------------------
    功能说明  : 抑制固定频率机械共振（丝杠固有频率、皮带拍频、伺服 300~800 Hz 尖叫）
                的带阻滤波；库内 LowPassFilter / HighPassFilter / SecondOrderFilter 都
                不带「中心频率 + Q 可调」的带阻形态，本件补该缺口；
                三道硬闸依次为：采样周期闸（决定采样频率，除零源头）、奈奎斯特闸
                （中心频率必须低于 0.45 倍采样频率，超了陷波会变成放大器）、
                系数分母闸（1 加 alpha 近零时拒绝重算并旁路）；
                参数在线改动只重算系数、保留历史状态不清零，避免改参瞬间断控制；
                输出双侧限幅并置饱和标志，是滤波发散前的最后一道防线。
    错误码    : 16#0002_2501 参数在线变更已重算系数（状态保留），或输出限幅生效——信息级，不置故障
                16#0002_2502 预留禁用（信息级，不得挪用）
                16#0002_2510 采样周期非法（不大于 0）——故障级，旁路输出
                16#0002_2511 中心频率超奈奎斯特 0.45 倍 / Q 越界 / 系数分母近零 / 限幅值非法——故障级，旁路输出
                16#0002_2512 预留禁用（故障级，不得挪用）
    码位总账  : 16#0002_2501 用 / 16#0002_2502 预留 ｜ 16#0002_2510 用 / 16#0002_2511 用 / 16#0002_2512 预留
    状态机    : 无 CASE，滤波状态由四个历史值承载，非法状态由参数闸拦截，不可能出现
    采样约定  : fbTrigReset 在本体首部无条件刷新；tSampleTime 必须等于本块所在任务的
                实际周期，否则中心频率与 Q 的物理含义失真，该参数不由本块测量。
    修订记录  : 2026-11-16 v1.0.0 首次入库（R18）
*)
FUNCTION_BLOCK FB_DL_NotchFilter
VAR_INPUT
    bEnable      : BOOL;                       // 使能，FALSE 时输出跟随输入并保持状态 / enable, FALSE passes the input through and keeps the state
    bReset       : BOOL;                       // 复位，上升沿清内部历史值 / reset, rising edge clears the internal history
    fIn          : REAL := 0.0;                // 输入信号，一般接位置或速度反馈 [用户单位] / input signal, usually a position or speed feedback [user unit]
    fCenterFreq  : REAL := 50.0;               // 陷波中心频率 [Hz]，范围 0.1~1000.0 / notch centre frequency [Hz], range 0.1~1000.0
    fQuality     : REAL := 2.0;                // 品质因数 Q [无量纲]，范围 0.1~50.0，越大陷波越窄 / quality factor Q [dimensionless], range 0.1~50.0, larger is narrower
    tSampleTime  : TIME := T#10MS;             // 采样周期 [ms]，范围 1~1000，必须等于任务周期 / sample period [ms], range 1~1000, must equal the task period
    fOutLimit    : REAL := 1.0E6;              // 输出幅值限幅，防系数病态发散 [用户单位]，必须大于 0 / output magnitude limit against ill-conditioned divergence [user unit], must exceed zero
END_VAR
VAR_OUTPUT
    fOut      : REAL;                          // 滤波输出 [用户单位] / filtered output [user unit]
    bSaturated: BOOL;                          // 输出被限幅（发散前兆）/ output clamped, a divergence precursor
    uCoeffRev : UDINT;                         // 系数重算次数，参数在线改动监视 [次] / coefficient recomputation count for online change monitoring [times]
    eErr      : UDINT;                         // 错误码，0=正常 / error id, 0=ok
    bError    : BOOL;                          // 故障标志，eErr 为故障级时 TRUE / error flag, TRUE on fault-level eErr
END_VAR
VAR
    fbTrigReset : R_TRIG;                      // 复位沿检测实例，本体首部无条件刷新 / reset edge instance, refreshed unconditionally
    fB0         : REAL;                        // 归一化分子系数 b0 [无量纲] / normalised numerator coefficient b0 [dimensionless]
    fB1         : REAL;                        // 归一化分子系数 b1 [无量纲] / normalised numerator coefficient b1 [dimensionless]
    fB2         : REAL;                        // 归一化分子系数 b2 [无量纲] / normalised numerator coefficient b2 [dimensionless]
    fA1         : REAL;                        // 归一化分母系数 a1 [无量纲] / normalised denominator coefficient a1 [dimensionless]
    fA2         : REAL;                        // 归一化分母系数 a2 [无量纲] / normalised denominator coefficient a2 [dimensionless]
    fA0         : REAL;                        // 分母基准，防零闸的被除数 [无量纲] / denominator base, the divisor under the zero gate [dimensionless]
    fX1         : REAL;                        // 输入历史值一 [用户单位] / input history one [user unit]
    fX2         : REAL;                        // 输入历史值二 [用户单位] / input history two [user unit]
    fY1         : REAL;                        // 输出历史值一 [用户单位] / output history one [user unit]
    fY2         : REAL;                        // 输出历史值二 [用户单位] / output history two [user unit]
    fOmega      : REAL;                        // 归一化角频率 [弧度] / normalised angular frequency [rad]
    fAlpha      : REAL;                        // 带宽系数 [无量纲] / bandwidth coefficient [dimensionless]
    fFs         : REAL;                        // 采样频率 [Hz] / sampling frequency [Hz]
    fCosW       : REAL;                        // 归一化角频率余弦，系数复用 [无量纲] / cosine of the normalised angular frequency, reused by the coefficients [dimensionless]
    fTs         : REAL;                        // 采样周期秒值 [s] / sample period in seconds [s]
    fPrevFc     : REAL;                        // 上一拍中心频率，变更检测 [Hz] / previous centre frequency for change detection [Hz]
    fPrevQ      : REAL;                        // 上一拍品质因数，变更检测 [无量纲] / previous quality factor for change detection [dimensionless]
    fPrevTs     : REAL;                        // 上一拍采样周期，变更检测 [s] / previous sample period for change detection [s]
    fY          : REAL;                        // 滤波结果中间量 [用户单位] / filter result intermediate [user unit]
    bInit       : BOOL := FALSE;               // 首扫标志，初值 FALSE，判据 NOT bInit / first-scan flag, initial FALSE, tested with NOT
    bParamBad   : BOOL;                        // 参数非法标志，本拍旁路 / parameter invalid flag, bypass this cycle
END_VAR
VAR CONSTANT
    DL_NOTCH_PI2      : REAL := 6.283185307;   // 二倍圆周率 [无量纲] / twice pi [dimensionless]
    DL_NOTCH_NYQ_RATIO: REAL := 0.45;          // 中心频率上限对采样频率的比值 [无量纲] / centre frequency cap as a fraction of the sampling frequency [dimensionless]
    DL_NOTCH_Q_MIN    : REAL := 0.1;           // Q 下限 [无量纲] / quality factor lower bound [dimensionless]
    DL_NOTCH_Q_MAX    : REAL := 50.0;          // Q 上限 [无量纲] / quality factor upper bound [dimensionless]
    DL_NOTCH_FC_MIN   : REAL := 0.1;           // 中心频率下限 [Hz] / centre frequency lower bound [Hz]
    DL_NOTCH_FC_MAX   : REAL := 1000.0;        // 中心频率上限 [Hz] / centre frequency upper bound [Hz]
    DL_NOTCH_TS_MAX   : REAL := 1.0;           // 采样周期上限秒值 [s] / sample period upper bound in seconds [s]
    DL_NOTCH_MS_SEC   : REAL := 1000.0;        // 毫秒转秒的除数，恒非零 [ms/s] / milliseconds to seconds divisor, never zero [ms/s]
    DL_NOTCH_TWO      : REAL := 2.0;           // 系数式中的常数二 [无量纲] / constant two in the coefficient formulas [dimensionless]
    DL_NOTCH_ONE      : REAL := 1.0;           // 系数式中的常数一 [无量纲] / constant one in the coefficient formulas [dimensionless]
    DL_NOTCH_CNT_MAX  : UDINT := 16#FFFF_FFFE; // 重算计数饱和值 [次] / recomputation counter saturation value [times]
    DL_FLOAT_EPS      : REAL := 1.0E-6;        // 浮点判等容差 [无量纲] / float equality tolerance [dimensionless]
    DL_NOTCH_INF_GUARD: REAL := 4.0E38;        // 非有限幅值判定阈值 [用户单位] / non-finite magnitude guard [user unit]
    DL_NOTCH_ZERO     : REAL := 0.0;           // 零值常量，避免裸字面量 [无量纲] / zero constant, avoids a bare literal [dimensionless]
END_VAR

// 段 1｜边沿实例无条件周期刷新（红线：严禁放入条件分支）/ segment 1, unconditional edge refresh
fbTrigReset(CLK := bReset);

// 段 2｜输出与错误状态预置 / segment 2, preset outputs and error status
eErr := 0;                                     // 预置无错误 / preset no error
bError := FALSE;                               // 预置无故障 / preset no fault
bSaturated := FALSE;                           // 预置未限幅 / preset not limited
bParamBad := FALSE;                            // 预置参数合法 / preset parameters valid

// 段 3｜首扫初始化（初值 FALSE，判据 NOT bInit）/ segment 3, first-scan initialisation
IF NOT bInit THEN
    fX1 := DL_NOTCH_ZERO;                      // 历史值清零 / clear the history
    fX2 := DL_NOTCH_ZERO;                      // 历史值清零 / clear the history
    fY1 := DL_NOTCH_ZERO;                      // 历史值清零 / clear the history
    fY2 := DL_NOTCH_ZERO;                      // 历史值清零 / clear the history
    uCoeffRev := 0;                            // 重算计数清零 / clear the recomputation counter
    fPrevFc := -DL_NOTCH_ONE;                  // 用不可能的值初始化，保证首拍必重算一次 / initialise with an impossible value so the first cycle always recomputes
    fPrevQ := -DL_NOTCH_ONE;                   // 同理用不可能值保证首拍必重算 / likewise impossible so first cycle recomputes
    fPrevTs := -DL_NOTCH_ONE;                  // 同理用不可能值保证首拍必重算 / likewise impossible so first cycle recomputes
    bInit := TRUE;                             // 首扫只做一次 / first scan runs once only
END_IF

// 段 4｜使能闸：失能即旁路且保持滤波状态 / segment 4, enable gate bypasses and keeps the state
IF NOT bEnable THEN
    fOut := fIn;                               // 输出跟随输入 / output follows the input
    RETURN;                                    // 失能即出口 / disabled is the exit
END_IF

// 段 5｜采样周期闸：决定采样频率，是全部除法的源头 / segment 5, sample period gate
IF tSampleTime <= T#0MS THEN
    eErr := 16#0002_2510;                      // 采样周期非法故障码 / illegal sample period fault id
    bError := TRUE;                            // 置故障标志 / raise the error flag
    fOut := fIn;                               // 旁路输出 / bypass the output
    RETURN;                                    // 故障级提前返回 / early return on fault
END_IF
fTs := TIME_TO_REAL(tSampleTime) / DL_NOTCH_MS_SEC; // 毫秒转秒 / milliseconds to seconds
IF (ABS(fTs) <= DL_FLOAT_EPS) OR (fTs > DL_NOTCH_TS_MAX) THEN
    eErr := 16#0002_2510;                      // 秒值近零或超上限，同属采样周期非法 / seconds near zero or above the cap, both are an illegal sample period
    bError := TRUE;                            // 置故障标志 / raise the error flag
    fOut := fIn;                               // 旁路输出 / bypass the output
    RETURN;                                    // 故障级提前返回 / early return on fault
END_IF

// 段 6｜奈奎斯特闸与 Q 域闸：超了陷波会变成放大器 / segment 6, Nyquist and quality factor gate
fFs := DL_NOTCH_ONE / fTs;                     // 采样频率，分母已过闸 / sampling frequency, the divisor already passed the gate
IF (fCenterFreq < DL_NOTCH_FC_MIN) OR (fCenterFreq > DL_NOTCH_FC_MAX) THEN
    eErr := 16#0002_2511;                      // 中心频率越界故障码 / centre frequency out of range fault id
    bError := TRUE;                            // 置故障标志 / raise the error flag
    bParamBad := TRUE;                         // 本拍旁路 / bypass this cycle
END_IF
IF fCenterFreq >= (DL_NOTCH_NYQ_RATIO * fFs) THEN
    eErr := 16#0002_2511;                      // 超奈奎斯特上限故障码 / above the Nyquist cap fault id
    bError := TRUE;                            // 置故障标志 / raise the error flag
    bParamBad := TRUE;                         // 本拍旁路 / bypass this cycle
END_IF
IF (fQuality < DL_NOTCH_Q_MIN) OR (fQuality > DL_NOTCH_Q_MAX) THEN
    eErr := 16#0002_2511;                      // Q 越界故障码 / quality factor out of range fault id
    bError := TRUE;                            // 置故障标志 / raise the error flag
    bParamBad := TRUE;                         // 本拍旁路 / bypass this cycle
END_IF
IF fOutLimit <= DL_FLOAT_EPS THEN
    eErr := 16#0002_2511;                      // 限幅值非法故障码（限幅失效等于失去发散保护）/ illegal limit fault id, a dead limit means no divergence protection
    bError := TRUE;                            // 置故障标志 / raise the error flag
    bParamBad := TRUE;                         // 本拍旁路 / bypass this cycle
END_IF
IF bParamBad THEN
    fOut := fIn;                               // 参数非法一律旁路 / any invalid parameter bypasses the filter
    RETURN;                                    // 故障级提前返回 / early return on fault
END_IF

// 段 7｜系数计算与分母防零闸 / segment 7, coefficient computation with the denominator guard
fOmega := DL_NOTCH_PI2 * fCenterFreq * fTs;    // 归一化角频率 / normalised angular frequency
fAlpha := SIN(fOmega) / (DL_NOTCH_TWO * fQuality); // 带宽系数，Q 已过闸恒非零 / bandwidth coefficient, the divisor is safe because Q passed the gate
fA0 := DL_NOTCH_ONE + fAlpha;                  // 分母基准 / denominator base
IF ABS(fA0) <= DL_FLOAT_EPS THEN
    eErr := 16#0002_2511;                      // 系数分母近零故障码 / coefficient denominator near zero fault id
    bError := TRUE;                            // 置故障标志 / raise the error flag
    fOut := fIn;                               // 旁路输出 / bypass the output
    RETURN;                                    // 故障级提前返回 / early return on fault
END_IF

// 段 8｜参数变更检测：变更只重算系数，历史状态保留不清零 / segment 8, parameter change detection keeps the state
IF (ABS(fCenterFreq - fPrevFc) > DL_FLOAT_EPS)
   OR (ABS(fQuality - fPrevQ) > DL_FLOAT_EPS)
   OR (ABS(fTs - fPrevTs) > DL_FLOAT_EPS) THEN
    fCosW := COS(fOmega);                      // 角频率余弦，四个系数共用 / cosine shared by the coefficients
    fB0 := DL_NOTCH_ONE / fA0;                 // 分子 b0，分母已过闸 / numerator b0, the divisor passed the gate
    fB1 := -DL_NOTCH_TWO * fCosW / fA0;        // 分子 b1 / numerator b1
    fB2 := fB0;                                // 分子 b2 与 b0 对称 / numerator b2 is symmetric to b0
    fA1 := -DL_NOTCH_TWO * fCosW / fA0;        // 分母 a1 / denominator a1
    fA2 := (DL_NOTCH_ONE - fAlpha) / fA0;      // 分母 a2 / denominator a2
    IF uCoeffRev < DL_NOTCH_CNT_MAX THEN
        uCoeffRev := uCoeffRev + 1;            // 饱和加一，绝不回绕 / saturating increment, never wraps
    END_IF
    eErr := 16#0002_2501;                      // 在线改参提示（信息级不置故障）/ online change hint, info level never raises a fault
    fPrevFc := fCenterFreq;                    // 记录中心频率 / remember the centre frequency
    fPrevQ := fQuality;                        // 记录品质因数 / remember the quality factor
    fPrevTs := fTs;                            // 记录采样周期 / remember the sample period
END_IF

// 段 9｜复位沿清状态（优先于滤波运算）/ segment 9, reset clears the history before filtering
IF fbTrigReset.Q THEN
    fX1 := DL_NOTCH_ZERO;                      // 历史值清零 / clear the history
    fX2 := DL_NOTCH_ZERO;                      // 历史值清零 / clear the history
    fY1 := DL_NOTCH_ZERO;                      // 历史值清零 / clear the history
    fY2 := DL_NOTCH_ZERO;                      // 历史值清零 / clear the history
END_IF

// 段 10｜直接 I 型二阶差分方程 / segment 10, direct form one second order difference equation
fY := fB0 * fIn + fB1 * fX1 + fB2 * fX2 - fA1 * fY1 - fA2 * fY2; // 二阶带阻 / second order band stop
IF (fY <> fY) OR (fY > DL_NOTCH_INF_GUARD) OR (fY < -DL_NOTCH_INF_GUARD) THEN
    fY := fY1;                                 // 非有限即退回上一拍输出，绝不让 NaN 进入状态 / non-finite falls back to the previous output, a NaN never enters the state
    bSaturated := TRUE;                        // 标记异常 / flag the anomaly
    eErr := 16#0002_2501;                      // 异常提示（信息级不置故障）/ anomaly hint, info level never raises a fault
END_IF

// 段 11｜输出双侧限幅 / segment 11, symmetrical output clamping
IF fY > fOutLimit THEN
    fY := fOutLimit;                           // 上侧限幅 / clamp the upper side
    bSaturated := TRUE;                        // 标记限幅 / flag the clamp
    eErr := 16#0002_2501;                      // 限幅提示（信息级不置故障）/ clamp hint, info level never raises a fault
ELSIF fY < -fOutLimit THEN
    fY := -fOutLimit;                          // 下侧限幅 / clamp the lower side
    bSaturated := TRUE;                        // 标记限幅 / flag the clamp
    eErr := 16#0002_2501;                      // 限幅提示（信息级不置故障）/ clamp hint, info level never raises a fault
END_IF

// 段 12｜状态推进与输出 / segment 12, push the state and publish the output
fX2 := fX1;                                    // 输入历史后移 / shift the input history
fX1 := fIn;                                    // 记录本拍输入 / record this cycle input
fY2 := fY1;                                    // 输出历史后移 / shift the output history
fY1 := fY;                                     // 记录本拍输出 / record this cycle output
fOut := fY;                                    // 对外输出 / publish the output
END_FUNCTION_BLOCK
